(* CODESYS project BODAS_RC18-12_27-18_40.library
   DocFormat: reStructuredText
   Company: Bosch Rexroth AG
   DefaultNamespace: BODAS_RC18-12_27-18_40
   Title: BODAS_RC18-12_27-18_40
   Description: User library to use BODAS-BSW services (API) for RC40.
   Version: 3.0.1

Project tree, tasks and I/O mapping:
  Communication API/
    CAN/
      STRUCTURE/
        data type bds_can_BufManage_ts
        data type bds_can_DataboxBufInfo_ts
        data type bds_can_DataboxData08_ts
        data type bds_can_Message_ts
        data type bds_can_DataboxData64_ts
        data type bds_can_RxDatabox_ts
        data type bds_can_DataboxData_ts
        data type bds_can_TxDatabox_ts
      ENUM/
        data type bds_can_Chnl_te
      CAN legacy/
        API/
          function bds_can_getData [ST]
          function bds_can_getDatabox [ST]
          function bds_can_getRxBufStatus [ST]
          function bds_can_getStatus [ST]
          function bds_can_getTxBufStatus [ST]
          function bds_can_init [ST]
          function bds_can_initRxDatabox [ST]
          function bds_can_initTxDatabox [ST]
          function bds_can_initxt [ST]
          function bds_can_isTxChannelFree [ST]
          function bds_can_isTxDataboxFree [ST]
          function bds_can_sendData [ST]
          function bds_can_sendDatabox [ST]
          function bds_can_registerBusOffCallback [ST]
          function bds_can_setTxDelay [ST]
          function bds_can_start [ST]
          function bds_can_resetTxBuf [ST]
          function bds_can_stop [ST]
          function bds_can_registerRxCallback [ST]
      CAN signal based/
        API/
          function bds_can_sendSignal [ST]
          function bds_can_sendSignalGroup [ST]
          function bds_can_receiveSignal [ST]
          function bds_can_receiveSignalGroup [ST]
          function bds_can_setGroupSignalData [ST]
          function bds_can_setMsgGroup [ST]
          function bds_can_resetAllMsgGroups [ST]
          function bds_can_startAllMsgGroups [ST]
      UNION/
        data type bds_can_DataboxData_tu
      GVL/
        global variables GVL_can
      CAN_FFI_API/
        function bds_can_sendData_ffi [ST]
        function bds_can_getData_ffi [ST]
        function bds_can_getStatus_ffi [ST]
        function bds_can_isTxChannelFree_ffi [ST]
        function bds_can_getRxBufStatus_ffi [ST]
        function bds_can_getTxBufStatus_ffi [ST]
        function bds_can_sendDatabox_ffi [ST]
        function bds_can_getDatabox_ffi [ST]
        function bds_can_isTxDataboxFree_ffi [ST]
      CAN-FD legacy/
        API/
          function bds_can_fd_getData [ST]
          function bds_can_fd_getRxBufStatus [ST]
          function bds_can_fd_getTxBufStatus [ST]
          function bds_can_fd_isTxChannelFree [ST]
          function bds_can_fd_registerRxBuf [ST]
          function bds_can_fd_registerTxBuf [ST]
          function bds_can_fd_resetTxBuf [ST]
          function bds_can_fd_sendData [ST]
          function bds_can_fd_registerRxCallback [ST]
          function bds_can_fd_registerRxDataboxes [ST]
          function bds_can_fd_registerTxDataboxes [ST]
          function bds_can_fd_initRxDatabox [ST]
          function bds_can_fd_initTxDatabox [ST]
          function bds_can_fd_getDatabox [ST]
          function bds_can_fd_sendDatabox [ST]
          function bds_can_fd_isTxDataboxFree [ST]
          function bds_can_fd_setTxDelay [ST]
        ENUM/
          data type bds_can_fd_St_te
        STRUCTURE/
          data type bds_can_fd_Message_ts
          data type bds_can_fd_RxDatabox_ts
          data type bds_can_fd_DataboxData_ts
          data type bds_can_fd_DataboxBufInfo_ts
          data type bds_can_fd_BufManage_ts
          data type bds_can_fd_TxDatabox_ts
      CAN_FD_FFI_API/
        function bds_can_fd_getRxBufStatus_ffi [ST]
        function bds_can_fd_sendData_ffi [ST]
        function bds_can_fd_getTxBufStatus_ffi [ST]
        function bds_can_fd_getData_ffi [ST]
        function bds_can_fd_isTxChannelFree_ffi [ST]
        function bds_can_fd_getDatabox_ffi [ST]
        function bds_can_fd_sendDatabox_ffi [ST]
        function bds_can_fd_isTxDataboxFree_ffi [ST]
    ISOBUS/
      STRUCTURE/
        data type bds_isobus_appInst_ts
        data type bds_isobus_bamCtrl_ts
        data type bds_isobus_caName_ts
        data type bds_isobus_canID_ts
        data type bds_isobus_dtcList_ts
        data type bds_isobus_dtc_ts
        data type bds_isobus_err_ts
        data type bds_isobus_rxDataboxInfo_ts
        data type bds_isobus_rxEtpCtrl_ts
        data type bds_isobus_rxMsg_ts
        data type bds_isobus_rxTpCtrl_ts
        data type bds_isobus_txDataboxInfo_ts
        data type bds_isobus_txEtpCtrl_ts
        data type bds_isobus_txMsg_ts
        data type bds_isobus_txTpCtrl_ts
        data type bds_isobus_lamp_ts
        data type bds_isobus_nm_ts
        data type bds_isobus_aperiodicDataboxNum_ts
        data type bds_isobus_periodicDataboxNum_ts
        data type bds_isobus_caAddrInfoTbl_ts
        data type bds_isobus_caAddrInfoTblRef_ts
      UNION/
        data type bds_isobus_caName_tu
        data type bds_isobus_canID_tu
      API/
        function bds_isobus_cfgAddrClaimFormat [ST]
        function bds_isobus_getCaAddr [ST]
        isobus dtclist bds_isobus_getDiagnostic [ST]
        function bds_isobus_getRxDataboxStatus [ST]
        function bds_isobus_getStatus [ST]
        function bds_isobus_initComm [ST]
        isobus dtclist bds_isobus_initDiagnostic [ST]
        function bds_isobus_registerErrClrCbk [ST]
        function bds_isobus_registerInstances [ST]
        function bds_isobus_registerRxDataboxes [ST]
        function bds_isobus_registerTxDataboxes [ST]
        function bds_isobus_sendDatabox [ST]
        function bds_isobus_sendRequestPGN [ST]
        function bds_isobus_setCaAddr [ST]
        function bds_isobus_setCaInfo [ST]
        function bds_isobus_setCaName [ST]
        function bds_isobus_initFailureList [ST]
        function bds_isobus_initRxDatabox [ST]
        function bds_isobus_initTxDatabox [ST]
        function bds_isobus_registerCaAddrTable [ST]
        function bds_isobus_registerCaAddrInfoCbk [ST]
        function bds_isobus_getCaAddrByName [ST]
        function bds_isobus_getAddressInfoTblRecordSize [ST]
      GVL/
        global variables GVL_isobus
      J1939-76/
        STRUCTURE/
          data type bds_isobus_cnsrDataboxInfo_ts
          data type bds_isobus_cnsrSdgMsg_ts
          data type bds_isobus_cnsrSdgSeqNum_ts
          data type bds_isobus_prodDataboxInfo_ts
          data type bds_isobus_prodSdgMsg_ts
          data type bds_isobus_sftyTmr_ts
          data type bds_isobus_sfty_canID_ts
          data type bds_isobus_shmMsg_ts
        API/
          function bds_isobus_initCnsrSdgDatabox [ST]
          function bds_isobus_initProdSdgDatabox [ST]
          function bds_isobus_registerCnsrSdgDataboxes [ST]
          function bds_isobus_registerProdSdgDataboxes [ST]
        UNION/
          data type bds_isobus_sdmCrcVal_tu
          data type bds_isobus_sfty_canID_tu
        ENUM/
          data type bds_isobus_sdgCnsrStatus_te
          data type bds_isobus_sdgState_te
          data type bds_isobus_sfty_apiRetVal_te
      ENUM/
        data type bds_isobus_caAddrCbEventType_te
    LIN/
      API/
        function bds_lin_getStatus [ST]
        function bds_lin_gotoSleep [ST]
        function bds_lin_receiveSignal [ST]
        function bds_lin_sendSignal [ST]
        function bds_lin_setSchedule [ST]
        function bds_lin_wakeUp [ST]
      GVL/
        global variables GVL_lin
    Ethernet/
      API/
        function bds_ethIPv4_setLocalIpAdr [ST]
        function bds_ethIPv4_getLocalIpAdr [ST]
        function bds_ethIPv4_setDoipAdr [ST]
        function bds_ethIPv4_getLinkState [ST]
      STRUCTURE/
        data type bds_ethIPv4_getLocalIpAdr_ts
        data type bds_ethIPv4_setLocalIpAdr_ts
        data type bds_ethIPv4_LocalIpAdr_ts
        data type bds_ethIPv4_linkStateInfo_ts
      ENUMS/
        data type bds_ethIPv4_statusApi_te
        data type bds_ethIPv4_linkState_te
        data type bds_ethIPv4_retDoipAdr_te
        data type bds_ethIPv4_retLinkState_te
  Diagnostics API/
    UDS/
      API/
        function bds_uds_disable [ST]
        function bds_uds_GetActiveDid [ST]
        function bds_uds_getActiveSession [ST]
        function bds_uds_getNodeID [ST]
        function bds_uds_permitAccess [ST]
        function bds_uds_registerDidReadCallback [ST]
        function bds_uds_registerDidWriteCallback [ST]
        function bds_uds_registerRoutineCtrlCallback [ST]
        function bds_uds_registerRoutineF000Callback [ST]
        function bds_uds_setCallbackStatus [ST]
        function bds_uds_setUUID [ST]
        function bds_uds_updNodeIDinNVM [ST]
        function bds_uds_registerEvalKeyCallback [ST]
        function bds_uds_registerGetSeedCallback [ST]
        function bds_uds_registerRoutineF001Callback [ST]
        Vehicle Identification Number(VIN) APIs/
          function bds_uds_setVin [ST]
          function bds_uds_getVin [ST]
          function bds_uds_registerVinCallback [ST]
        function bds_uds_getActiveService [ST]
        function bds_uds_setNodeIdTesterId [ST]
      UNION/
        data type bds_uds_udsconfigparameter_tu
      STRUCTURE/
        data type bds_uds_udsconfigparameter_ts
        data type bds_uds_getActiveService_ts
      GVL/
        global variables GVL_uds
      FFI_API/
        function bds_uds_getActiveSession_ffi [ST]
        function bds_uds_getNodeID_ffi [ST]
        function bds_uds_getActiveService_ffi [ST]
        function bds_uds_getActiveDid_ffi [ST]
      ENUM/
        data type bds_udsCmn_statusApi_te
        data type bds_uds_setNodeIdTesterId_te
    XCP/
      API/
        function bds_xcp_setMode [ST]
      GVL/
        global variables GVL_xcp
  I/O API/
    SAFOUT/
      STRUCTURE/
        data type bds_safout_ts
      API/
        function bds_safout_resetError [ST]
        function bds_safout_ignoreError [ST]
        function bds_safout_getStatus [ST]
        function bds_safout_unlock [ST]
        function bds_safout [ST]
        function bds_safout_cfg [ST]
        function bds_safout_cfgDiag [ST]
        function bds_safout_enableTest [ST]
      GVL/
        global variables GVL_safout
    IN legacy/
      STRUCTURE/
        data type bds_in_aic_ts
        data type bds_in_fi_ts
        data type bds_in_FrqBuffered_ts
        data type bds_in_aiv_ts
        data type bds_in_sent_SDDataBox_ts
        data type bds_in_sent_slowData_ts
        data type bds_in_stPhase_ts
        data type bds_in_ri_ts
        data type bds_in_sent_BufManage_ts
        data type bds_in_sent_copyFDBuf_ts
        data type bds_in_sent_databoxinfo_ts
        data type bds_in_sent_decodedFD_ts
        data type bds_in_sent_FDBufInfo_ts
        data type bds_in_phase_ts
      API/
        function bds_in_aic_getStatus [ST]
        function bds_in_aid [ST]
        function bds_in_aid_cfg [ST]
        function bds_in_aiv [ST]
        function bds_in_aiv_cfg [ST]
        function bds_in_phase [ST]
        function bds_in_fi_cfg [ST]
        function bds_in_fi_getStatus [ST]
        function bds_in_phase_getStatus [ST]
        function bds_in_phase_resetCounter [ST]
        function bds_in_ri_cfg [ST]
        function bds_in_ri_cfgTemp [ST]
        function bds_in_sent_getSDDatabox [ST]
        function bds_in_sent_getStatus [ST]
        function bds_in_sent_initSDDatabox [ST]
        function bds_in_sent_registerCopyFDFifo [ST]
        function bds_in_sent_registerFDFifo [ST]
        function bds_in_ri_getStatus [ST]
        function bds_in_aiv_getStatus [ST]
        function bds_in_sent_registerSDDataboxes [ST]
        function bds_in_sent_getSD [ST]
        function bds_in_ri [ST]
        function bds_in_ai [ST]
        function bds_in_aic [ST]
        function bds_in_ri_getTemp [ST]
        function bds_in_sent_copyFDFifo [ST]
        function bds_in_sent_disable [ST]
        function bds_in_sent_enable [ST]
        function bds_in_sent_getFD [ST]
        function bds_in_aic_cfg [ST]
        function bds_in_di [ST]
        function bds_in_fi [ST]
        function bds_in_fi_buffered [ST]
      GVL/
        global variables GVL_in
    OUT_LEGACY/
      function bds_out_do_resetError [ST]
      function bds_out_do_unlock [ST]
      function bds_out_po [ST]
      function bds_out_poc [ST]
      function bds_out_poc_cfgDither [ST]
      function bds_out_poc_cfgPI [ST]
      function bds_out_po_cfgPwrLs [ST]
      function bds_out_po_cfg [ST]
      function bds_out_po_disableTstPls [ST]
      function bds_out_po_getCurrent [ST]
      function bds_out_po_getStatus [ST]
      function bds_out_po_resetError [ST]
      function bds_out_po_cfgPeriod [ST]
      function bds_out_po_disable [ST]
      function bds_out_aov_cfg [ST]
      function bds_out_aov_cfgPI [ST]
      function bds_out_aov_getStatus [ST]
      function bds_out_aov_getVoltage [ST]
      function bds_out_aov_resetError [ST]
      function bds_out_cfgLoadCharacteristic [ST]
      function bds_out_do [ST]
      function bds_out_do_cfgPwrLs [ST]
      function bds_out_do_disable [ST]
      function bds_out_aov [ST]
      function bds_out_do_disableTstPls [ST]
      function bds_out_do_getCurrent [ST]
      function bds_out_pod [ST]
      function bds_out_do_getStatus [ST]
      function bds_out_poc_cfg [ST]
      function bds_out_po_unlock [ST]
    OUT/
      API/
        function bds_outClcU_setVoltage [ST]
        function bds_outClcU_setPercUBat [ST]
        function bds_outClcU_get [ST]
        function bds_outClcU_rstErr [ST]
        function bds_outDig_set [ST]
        function bds_outDig_get [ST]
        function bds_outDig_cfgDiag [ST]
        function bds_outDig_rstErr [ST]
        function bds_outPwm_setDutyCycle [ST]
        function bds_outPwm_get [ST]
        function bds_outPwm_cfgPeriod [ST]
        function bds_outPwm_rstErr [ST]
        function bds_outPwm_cfgDiag [ST]
        function bds_outPwm_cfgMode [ST]
        function bds_outPwm_setCurrent [ST]
        function bds_outPwm_cfgDiagCurrentDe [ST]
        function bds_outPwm_cfgClc [ST]
        function bds_outPwm_cfgDither [ST]
        function bds_outClcU_cfgClc [ST]
      STRUCTURE/
        data type bds_out_do_ts
        data type bds_out_po_ts
        data type bds_out_aov_ts
        data type bds_outClcU_setVoltage_ts
        data type bds_outClcU_setPercUBat_ts
        data type bds_outClcU_get_ts
        data type bds_outCmn_statusDiag_tb
        data type bds_outClcU_rstErr_ts
        data type bds_outDig_set_ts
        data type bds_outDig_get_ts
        data type bds_outDig_cfgDiag_ts
        data type bds_outDig_rstErr_ts
        data type bds_outPwm_setDutyCycle_ts
        data type bds_outPwm_get_ts
        data type bds_outPwm_cfgPeriod_ts
        data type bds_outPwm_rstErr_ts
        data type bds_outPwm_cfgDiag_ts
        data type bds_outPwm_cfgMode_ts
        data type bds_outPwm_setCurrent_ts
        data type bds_outPwm_cfgDiagCurrentDe_ts
        data type bds_outPwm_cfgDither_ts
        data type bds_outClcU_cfgClc_ts
        data type bds_outClcU_clcParams_ts
        data type bds_outCmn_diagParam_ts
        data type bds_outPwm_cfgClc_ts
        data type bds_outPwm_clcParams_ts
        data type bds_outPwm_ditherParams_ts
      ENUM/
        data type bds_load_characteristic_te
        data type bds_outCmn_statusApi_te
        data type bds_outPwm_cfgMode_te
        data type bds_outPwm_cfgDither_te
      GVL/
        global variables GVL_out
      FFI_API/
        function bds_out_aov_ffi [ST]
        function bds_out_aov_cfg_ffi [ST]
        function bds_out_aov_cfgPI_ffi [ST]
        function bds_out_aov_getStatus_ffi [ST]
        function bds_out_aov_getVoltage_ffi [ST]
        function bds_out_cfgLoadCharacteristic_ffi [ST]
        function bds_out_do_ffi [ST]
        function bds_out_do_cfgPwrLs_ffi [ST]
        function bds_out_do_disable_ffi [ST]
        function bds_out_do_disableTstPls_ffi [ST]
        function bds_out_do_getCurrent_ffi [ST]
        function bds_out_do_getStatus_ffi [ST]
        function bds_out_po_ffi [ST]
        function bds_out_poc_ffi [ST]
        function bds_out_poc_cfg_ffi [ST]
        function bds_out_poc_cfgDither_ffi [ST]
        function bds_out_poc_cfgPI_ffi [ST]
        function bds_out_pod_ffi [ST]
        function bds_out_po_cfg_ffi [ST]
        function bds_out_po_cfgPeriod_ffi [ST]
        function bds_out_po_cfgPwrLs_ffi [ST]
        function bds_out_po_disable_ffi [ST]
        function bds_out_po_disableTstPls_ffi [ST]
        function bds_out_po_getCurrent_ffi [ST]
        function bds_out_po_getStatus_ffi [ST]
    SENT/
      STRUCTURE/
        data type bds_sent_chSt_tb
        data type bds_sent_rxFastData_ts
        data type bds_sent_rxSlowData_ts
        data type bds_sent_getSlowDataBufd_ts
        data type bds_sent_getFastDataBufd_ts
        data type bds_sent_fastDataMsg_ts
        data type bds_sent_fastDataBuf_ts
        data type bds_sent_slowDataMsg_ts
        data type bds_sent_slowDataBuf_ts
      ENUM/
        data type bds_sentCmn_status_te
      API/
        function bds_sent_getFastData [ST]
        function bds_sent_getSlowData [ST]
        function bds_sent_getFastDataBufd [ST]
        function bds_sent_getSlowDataBufd [ST]
      FFI_API/
        function bds_sent_getFastData_ffi [ST]
        function bds_sent_getFastDataBufd_ffi [ST]
        function bds_sent_getSlowData_ffi [ST]
        function bds_sent_getSlowDataBufd_ffi [ST]
    IN/
      STRUCTURE/
        data type bds_inI_measmt_ts
        data type bds_inDig_measmt_ts
        data type bds_inCmn_pullParam_ts
        data type bds_inI_cfgPull_ts
        data type bds_inI_shunt_ts
        data type bds_inDig_cfgPull_ts
        data type bds_inPwm_tiMeasmt_ts
        data type bds_inPwm_tiBufdMeasmt_ts
        data type bds_inPwm_frqMeasmt_ts
        data type bds_inPwm_tiBufd_ts
        data type bds_inR_measmt_ts
        data type bds_inU_measmt_ts
        data type bds_inU_cfgPull_ts
        data type bds_inPha_measmt_ts
        data type bds_inPha_statusDiag_tb
        data type bds_inPha_tiBufdMeasmt_ts
        data type bds_inPha_tiBufd_ts
      ENUM/
        data type bds_inCmn_status_te
        data type bds_inCmn_pullType_te
        data type bds_inI_stShunt_te
        data type bds_inCmn_iPull_te
      API/
        function bds_inI_cfgPull [ST]
        function bds_inI_ctrlShunt [ST]
        function bds_inDig_get [ST]
        function bds_inI_get [ST]
        function bds_inDig_cfgPull [ST]
        function bds_inPwm_getTi [ST]
        function bds_inPwm_getTiBufd [ST]
        function bds_inR_get [ST]
        function bds_inPwm_getFrq [ST]
        function bds_inU_get [ST]
        function bds_inU_cfgPull [ST]
        function bds_inPha_get [ST]
        function bds_inPha_getTiBufd [ST]
      FFI_API/
        function bds_inDig_cfgPull_ffi [ST]
        function bds_inI_cfgPull_ffi [ST]
        function bds_inI_ctrlShunt_ffi [ST]
        function bds_inPwm_getFrq_ffi [ST]
        function bds_inPwm_getTi_ffi [ST]
        function bds_inPwm_getTiBufd_ffi [ST]
        function bds_inU_cfgPull_ffi [ST]
  Memory API/
    NVM/
      API/
        function bds_mem_getBlockStatus [ST]
        function bds_mem_markBlock [ST]
        function bds_mem_readBlock [ST]
        function bds_mem_writeBlock [ST]
      GVL/
        global variables GVL_mem
      FFI_API/
        function bds_mem_getBlockStatus_ffi [ST]
        function bds_mem_markBlock_ffi [ST]
        function bds_mem_readBlock_ffi [ST]
        function bds_mem_writeBlock_ffi [ST]
  System API/
    SEC/
      ENUM/
        data type bds_diag_inst_te
        data type bds_sec_securityOperations_te
      API/
        function bds_sec_evalRespKey [ST]
        function bds_sec_getLevel [ST]
        function bds_sec_getRnd [ST]
        function bds_sec_resetLevel [ST]
        function bds_sec_saveSecret [ST]
        function bds_sec_scrambleRexrothSecretsPerm [ST]
        function bds_sec_setLevel [ST]
        function bds_sec_getSeed [ST]
      GVL/
        global variables GVL_sec
    SYS/
      API/
        function bds_sys_ait [ST]
        function bds_sys_aiv [ST]
        function bds_sys_cancelAltWakeup [ST]
        function bds_sys_di [ST]
        function bds_sys_do [ST]
        function bds_sys_getAge [ST]
        function bds_sys_getCoreLoad [ST]
        function bds_sys_getEcuInfo [ST]
        function bds_sys_getResetInfo [ST]
        function bds_sys_getStates [ST]
        function bds_sys_getT15 [ST]
        function bds_sys_getTaskRuntime [ST]
        function bds_sys_getTime [ST]
        function bds_sys_getVersion [ST]
        function bds_sys_getVSS [ST]
        function BDS_SYS_GET_LOCK_COMMON [ST]
        function bds_sys_memByteCopy [ST]
        function bds_sys_releasePostRunProlong [ST]
        function BDS_SYS_RELEASE_LOCK_COMMON [ST]
        function bds_sys_requestPostRunProlong [ST]
        function bds_sys_resetCoreLoad [ST]
        function bds_sys_resetEcu [ST]
        function bds_sys_resetINH [ST]
        function bds_sys_setVSS [ST]
        function bds_sys_startLoader [ST]
        function bds_sysPb_getVariant [ST]
        function bds_sysPb_cfgVariant [ST]
        function bds_sys_applSwName [ST]
        function bds_sysSm_getCfg [ST]
        function bds_sys_regOverwriteOpHrsCbk [ST]
        function bds_codesys_setForcingWritingMode [ST]
      ENUM/
        data type bds_sys_coreid_te
        data type bds_sys_states_te
        data type bds_sys_task_te
        data type bds_sysCmn_status_te
        data type bds_sys_aswNameStatus_te
        data type bds_sys_regOverwriteOpHrs_te
      STRUCTURE/
        data type bds_sys_coreload_info_ts
        data type bds_sys_states_ts
        data type bds_sys_taskruntime_ts
        data type bds_ResetInfo_ts
        data type bds_EcuInfo_ts
        data type bds_sysPb_retValCfgVrnt_ts
        data type bds_sysPb_vrntParam_ts
        data type bds_sysPb_retValGetVrnt_ts
        data type bds_sys_retValApplSwName_ts
      GVL/
        global variables GVL_sys
      FFI_API/
        function bds_sysPb_getVariant_ffi [ST]
        function bds_sys_getAge_ffi [ST]
        function bds_sys_getCoreLoad_ffi [ST]
        function bds_sys_getEcuInfo_ffi [ST]
        function bds_sys_getResetInfo_ffi [ST]
        function bds_sys_getStates_ffi [ST]
        function bds_sys_getTaskRuntime_ffi [ST]
        function bds_sys_getTime_ffi [ST]
        function bds_sys_getVersion_ffi [ST]
    DSM/
      STRUCTURE/
        data type bds_dfes_ts
        data type bds_dsm_j1939Lamp_ts
        data type bds_dsm_J1939_info_ts
        data type bds_dsm_dfc_ts
        data type bds_dsm_dtcj1939_ts
        data type bds_dsm_fid_ts
      API/
        function bds_dsm_delError [ST]
        function bds_dsm_delErrors [ST]
        function bds_dsm_delErrorsJ1939 [ST]
        function bds_dsm_delError_DTC [ST]
        Macro Functions/
          function bds_dsm_DFC_da [ST]
          function bds_dsm_DFC_dfl [ST]
          function bds_dsm_DFC_fl [ST]
          function bds_dsm_DFC_fsc [ST]
          function bds_dsm_DFC_ldf [ST]
          function bds_dsm_DFC_ms [ST]
          function bds_dsm_DFC_t [ST]
          function bds_dsm_DFC_tf [ST]
          function bds_dsm_DFC_tsc [ST]
        function bds_dsm_getErrors [ST]
        function bds_dsm_getDTC_Status [ST]
        function bds_dsm_getErrors_DTC [ST]
        function bds_dsm_getFIdPermission [ST]
        function bds_dsm_getNumErrors [ST]
        function bds_dsm_getNumErrorsJ1939 [ST]
        function bds_dsm_testError [ST]
        function bds_dsm_test_ErrorDFC [ST]
        function bds_dsm_test_ErrorDTC [ST]
        function bds_dsm_updateDebError [ST]
        function bds_dsm_updateError [ST]
        function bds_dsm_updateError_DTC [ST]
        function bds_dsm_getDFC_Status [ST]
        function bds_dsm_getDFES [ST]
        function bds_dsm_getErrorsJ1939 [ST]
        function bds_dsm_getDFES_DTC [ST]
        function bds_dsm_getDTC_DFC [ST]
        function bds_dsm_getDTC_DFCJ1939 [ST]
        function bds_dsm_getDTC_J1939 [ST]
      ENUM/
        data type bds_dsm_state_te
      GVL/
        global variables GVL_dsm
      FFI_API/
        function bds_dsm_getErrors_ffi [ST]
        function bds_dsm_updateError_ffi [ST]
        function bds_dsm_getNumErrors_ffi [ST]
        function bds_dsm_getDFC_Status_ffi [ST]
      DSM Refactored( 3-byte DTC)/
        STRUCTURE/
          data type bds_dsmCmn_stWord_tb
          data type bds_dsmDTC_deleteErr_ts
          data type bds_dsmDTC_getDFES_ts
          data type bds_dsmDTC_getDTCVal_ts
          data type bds_dsmDTC_getErrList_ts
          data type bds_dsmDTC_getStatus_ts
          data type bds_dsmDTC_updateErr_ts
          data type bds_dsmJ1939_LampSt_tb
          data type bds_dsmJ1939_getJ1939DTC_ts
        API/
          function bds_dsmDTC_getDTCVal [ST]
          function bds_dsmDTC_updateErr [ST]
          function bds_dsmDTC_deleteErr [ST]
          function bds_dsmDTC_getErrList [ST]
          function bds_dsmDTC_getStatus [ST]
          function bds_dsmDTC_getDFES [ST]
          function bds_dsmJ1939_getJ1939DTC [ST]
        ENUM/
          data type bds_dsmCmn_st_te
          data type bds_dsmCmn_errState_te
          data type bds_dsmCmn_fltLvl_te
*)

// Communication API/CAN/STRUCTURE/bds_can_BufManage_ts
{attribute 'external_name' := 'cmp_rts_bds_can_BufManage_ts'}
TYPE bds_can_BufManage_ts :
STRUCT
	length_u16: UINT;
	idx_in_u16: UINT;
	idx_out_u16: UINT;
	BufEmpty_l: BOOL;
	BufOvfl_l: BOOL;
END_STRUCT
END_TYPE

// Communication API/CAN/ENUM/bds_can_Chnl_te
{attribute 'external_name' := 'cmp_rts_bds_can_Chnl_te'}
TYPE bds_can_Chnl_te :
(
	///CAN channel 1
	BDS_CAN_1_D := 0,
	///CAN channel 2
	BDS_CAN_2_D,
	///CAN channel 3
	BDS_CAN_3_D,
	///CAN channel 4
	BDS_CAN_4_D,
	BDS_CAN_NBR_E
)USINT;
END_TYPE

// Communication API/CAN/STRUCTURE/bds_can_DataboxBufInfo_ts
{attribute 'external_name' := 'cmp_rts_bds_can_DataboxBufInfo_ts'}
TYPE bds_can_DataboxBufInfo_ts :
STRUCT
	start_pas: POINTER TO bds_can_DataboxData_ts;
	Manage_s: bds_can_BufManage_ts;
END_STRUCT
END_TYPE

// Communication API/CAN/STRUCTURE/bds_can_DataboxData08_ts
{attribute 'external_name' := 'cmp_rts_bds_can_DataboxData08_ts'}
TYPE bds_can_DataboxData08_ts :
STRUCT
	data_au8: ARRAY[0..7] OF USINT;
	numBytes_u8: USINT;
END_STRUCT
END_TYPE

// Communication API/CAN/UNION/bds_can_DataboxData_tu
{attribute 'external_name' := 'cmp_rts_bds_can_DataboxData_tu'}
TYPE bds_can_DataboxData_tu :

UNION
	len08_s: bds_can_DataboxData08_ts;
	len64_s: bds_can_DataboxData64_ts;
END_UNION

END_TYPE

// Communication API/CAN/STRUCTURE/bds_can_Message_ts
{attribute 'external_name' := 'cmp_rts_bds_can_Message_ts'}
TYPE bds_can_Message_ts :
STRUCT
	///Identifier of the message.
	id_u32: UDINT;
	///Format which will be transmitted (Standard / Extended)
	format_u8: USINT;
	///Number of data bytes which will be transmitted or which where received.
	numBytes_u8: USINT;
	///Data which will be transmitted or which were received.
	data_au8: ARRAY[0..7] OF USINT;
END_STRUCT
END_TYPE

// Communication API/CAN/STRUCTURE/bds_can_DataboxData64_ts
{attribute 'external_name' := 'cmp_rts_bds_can_DataboxData64_ts'}
TYPE bds_can_DataboxData64_ts :
STRUCT
	data_au8: ARRAY[0..63] OF USINT;
	numBytes_u8: USINT;
END_STRUCT
END_TYPE

// Communication API/CAN/STRUCTURE/bds_can_RxDatabox_ts
{attribute 'external_name' := 'cmp_rts_bds_can_RxDatabox_ts'}
TYPE bds_can_RxDatabox_ts :
STRUCT
	id_u32: UDINT;
	format_u8: USINT;
	numBytes_u8: USINT;
	callback_pf: UDINT;
	Buf_s: bds_can_DataboxBufInfo_ts;
END_STRUCT
END_TYPE

// Communication API/CAN/STRUCTURE/bds_can_DataboxData_ts
{attribute 'external_name' := 'cmp_rts_bds_can_DataboxData_ts'}
TYPE bds_can_DataboxData_ts :
STRUCT
	///Data which will be transmitted or which were received.
	data_au8: ARRAY[0..7] OF USINT;
	///Number of data bytes which will be transmitted or which where received.
	numBytes_u8: USINT;
END_STRUCT
END_TYPE

// System API/DSM/STRUCTURE/bds_dfes_ts
{attribute 'external_name' := 'cmp_rts_bds_dfes_ts'}
TYPE bds_dfes_ts :
STRUCT
	/// REFERENCE number
	id: UINT := 12;
	/// assigned predebouncing mode
	debmode: UINT := 4;
END_STRUCT
END_TYPE

// System API/SEC/ENUM/bds_diag_inst_te
{attribute 'external_name' := 'cmp_rts_bds_diag_inst_te'}
TYPE bds_diag_inst_te :
(
	BDS_SEC_ASW_START_INSTANCE_E := 0,
	BDS_SEC_ASW_INST_NAME_1_E := BDS_SEC_ASW_START_INSTANCE_E,
	BDS_SEC_ASW_INST_NAME_2_E,
	BDS_SEC_ASW_INST_NAME_3_E,
	BDS_SEC_ASW_NUM_INSTANCE_E
);
END_TYPE

// I/O API/OUT/STRUCTURE/bds_out_do_ts
{attribute 'external_name' := 'cmp_rts_bds_out_do_ts'}
TYPE bds_out_do_ts :
STRUCT
	///status flags for status_b16 
	///	initOut_DB16: USINT := 16#1;(*initialization after startup*)
	///	
	///	cfgPOC_DB16: USINT := 16#2;(*configuration of closed loop control*)
	///	
	///	cfgPeriod_DB16: USINT := 16#4;(*configuration of period*)
	///	
	///	cfgDither_DB16: USINT := 16#8;(*configuration of dither*)
	///	
	///	cfgDeviation_DB16: USINT := 16#10;(*configuration of deviation*)
	///	
	///	cfgPI_DB16: USINT := 16#20;(*configuration of KpKi*)
	///	
	///	lockedSCB_DB16: USINT := 16#40;(*locked by SCB...necessary for AOV*)
	///	
	///	lockedSCG_DB16: USINT := 16#80;(*locked by SCG...necessary for AOV*)
	///	
	///	lockedOC_DB16: UINT := 16#100;(*locked by OC*)
	///	
	///	locked_DB16: UINT := 16#200;(*locked by Error Handler*)
	///	
	///	lockedMO_DB16: UINT := 16#400;(*locked by Monitoring Module (MO) Error*)
	///	
	///	lockCouTiReact_DB16: UINT := 16#800;(*locked reactivation timer reload after a hot short circuit*)
	///	
	///	tiReactNotElapsed_DB16: UINT := 16#1000;(*time for reactivation after a hot short circuit not elapsed*)
	///	
	///	linked_DB16: UINT := 16#2000;(*linked at least with one other safout output*)
	///	
	///	tlsPlsDis_DB16: UINT:=16#4000;(*Test pulses disable*)
	///	
	///	disabled_DB16: UINT := 16#8000;(*output is disabled (avoid open load faults of unused outputs)*)
	///	
	///	cfgOutMask_DB16: UINT := ((((cfgPI_DB16 OR cfgDeviation_DB16) OR cfgDither_DB16) OR cfgPeriod_DB16) OR cfgPOC_DB16);
	status_b16: UINT;
	///state
	state_u8: USINT;
	///ADC digits, range from 0..25000
	digits_u16: UINT;
	///actual current [mA]
	iAct_u16: UINT;
	///fault status
	stDFC_SCB_u16: UINT;
	///fault status
	stDFC_SCG_u16: UINT;
	///fault status
	stDFC_OL_u16: UINT;
	///fault status
	stDFC_OT_u16: UINT;
	///fault status
	stDFC_OC_u16: UINT;
	///Unintended switch ON of output
	unintendedSwitchONErr_l: BOOL;
	///locked by Inhibits
	lockedByINH_l: BOOL;
END_STRUCT
END_TYPE

// I/O API/IN legacy/STRUCTURE/bds_in_aic_ts
{attribute 'external_name' := 'cmp_rts_bds_in_aic_ts'}
TYPE bds_in_aic_ts :
STRUCT
	///status flags for status_b16 
	///	
	///	initIn_DB16: USINT := 16#1;(*initialization after startup*)
	///	
	///	cfgAiv_DB16: USINT := 16#2;(*configured for AIV thresholds*)
	///	
	///	cfgAic_DB16: USINT := 16#4;(*configured for AIC thresholds*)
	///	
	///	cfgAid_DB16: USINT := 16#8;(*configured for AID thresholds*)
	///	
	///	cfgRi_DB16: USINT := 16#10;(*configured for RI thresholds*)
	///	
	///	cfgFreq_DB16: USINT := 16#20;(*configured for standard frequency sensor*)
	///	
	///	cfgFreqDSM_DB16: USINT := 16#40;(*configured for DSM frequency sensor*)
	///	
	///	lostSignalInfoDSM_DB16: USINT := 16#80;
	///	
	///	actShunt_DB16: UINT := 16#1000;(*shunt is activated for DSM sensor respective AIC*)
	///	
	///	lockReactShunt_DB16: UINT := 16#2000;(*locked shunt reactivation*)
	///	
	///	cfgInMask_DB16: UINT := (((((cfgFreqDSM_DB16 OR cfgFreq_DB16) OR cfgRi_DB16) OR cfgAid_DB16) OR cfgAic_DB16) OR cfgAiv_DB16);
	status_b16: UINT;
	///ADC digits, range from 0..25000
	digits_u16: UINT;
	///current [µA]
	i_uA_u16: UINT;
	///fault status
	stDFC_SCB_u16: UINT;
	///fault status
	stDFC_SCG_u16: UINT;
END_STRUCT
END_TYPE

// I/O API/IN legacy/STRUCTURE/bds_in_fi_ts
{attribute 'external_name' := 'cmp_rts_bds_in_fi_ts'}
TYPE bds_in_fi_ts :
STRUCT
	///status flags for status_b16 
	///	
	///	initIn_DB16: USINT := 16#1;(*initialization after startup*)
	///	
	///	cfgAiv_DB16: USINT := 16#2;(*configured for AIV thresholds*)
	///	
	///	cfgAic_DB16: USINT := 16#4;(*configured for AIC thresholds*)
	///	
	///	cfgAid_DB16: USINT := 16#8;(*configured for AID thresholds*)
	///	
	///	cfgRi_DB16: USINT := 16#10;(*configured for RI thresholds*)
	///	
	///	cfgFreq_DB16: USINT := 16#20;(*configured for standard frequency sensor*)
	///	
	///	cfgFreqDSM_DB16: USINT := 16#40;(*configured for DSM frequency sensor*)
	///	
	///	lostSignalInfoDSM_DB16: USINT := 16#80;
	///	
	///	actShunt_DB16: UINT := 16#1000;(*shunt is activated for DSM sensor respective AIC*)
	///	
	///	lockReactShunt_DB16: UINT := 16#2000;(*locked shunt reactivation*)
	///	
	///	cfgInMask_DB16: UINT := (((((cfgFreqDSM_DB16 OR cfgFreq_DB16) OR cfgRi_DB16) OR cfgAid_DB16) OR cfgAic_DB16) OR cfgAiv_DB16);
	///	
	///	standstill_DU8: USINT := 16#0;(*standstill*)
	///	
	///	dirLeft_DU8: USINT := 16#1;(*direction left*)
	///	
	///	dirRight_DU8: USINT := 16#2;(*direction right*)
	///	
	///	dirUnknown_DU8: USINT := 16#4;(*direction not known for sure (e.g. after standstill)*)
	///	
	///	noError_DU8: USINT := 16#0;(*error free*)
	///	
	///	airGapError_DU8: USINT := 16#1;(*air gap error (pulse is shorter than 64us)*)
	///	
	///	mountError_DU8: USINT := 16#2;(*mounting error (pulse is longer than 254us)*)
	///	
	///	signalLengthError_DU8: USINT := 16#4;(*undefined signal length - should not occur (pulse is longer than 1785us*)
	///	
	///	signalError_DU8: USINT := 16#8;(*period too long or measured period exceeds maximum period*)
	///	
	///	noStatusAvailable_DU8: USINT := 16#10;(*no status signal available (frequency to high)*)
	///	
	///	diagSCUBAT_DU8: USINT := 16#20;
	///	
	///	diagSCGND_OR_OL_DU8: USINT := 16#40;
	///	
	///	maskFrequency_DU32: UDINT := 16#FFFFF;(*DSM mask to get the frequency out*)
	///	
	///	maskDirection_DU32: UDINT := 16#F00000;(*DSM mask to get the direction*)
	///	
	///	numShiftDirection_DU32: USINT := 20;(*DSM shift number to get the direction*)
	///	
	///	maskStatus_DU32: UDINT := 16#FF000000;(*DSM mask to get the status*)
	///	
	///	numShiftStatus_DU32: USINT := 24;(*DSM shift number to get the status*)
	status_b16: UINT;
	///current dutycycle [100%=16#8000]
	rDutycycle_u32: UDINT;
	///last high_time duration [µs]
	tiPulse_u32: UDINT;
	///period duration [µs]
	tiPeriod_u32: UDINT;
	///signal period counter
	ctPeriod_u32: UDINT;
	///signal state
	///   + Bit0 state at function call time ("1" for high or "0" for low
	///   + Bit1 no update available (request within the same period)
	///   + Bit2 period too long (timer overflow)
	///   + Bit3 measured period exceeds given maximum length 
	stSignal_u8: USINT;
	///frequency in [dHz]
	f_dHz_u32: UDINT;
	///period duration [µs] for DSM sensor
	tiPeriodDSM_u32: UDINT;
	///frequency of DSM in [dHz] (see defines above)
	f_dHzDSM_u32: UDINT;
	///direction (see defines above)
	directionDSM_u8: USINT;
	///status
	statusDSM_u8: USINT;
END_STRUCT
END_TYPE

// I/O API/IN legacy/STRUCTURE/bds_in_FrqBuffered_ts
{attribute 'external_name' := 'cmp_rts_bds_in_FrqBuffered_ts'}
TYPE bds_in_FrqBuffered_ts :
STRUCT
	///Pointer of the start address of the period array
	tiPeriod_pu32: POINTER TO UDINT;
	///Pointer of the start address of the pulse array
	tiPulse_pu32: POINTER TO UDINT;
END_STRUCT
END_TYPE

// Communication API/CAN/STRUCTURE/bds_can_TxDatabox_ts
{attribute 'external_name' := 'cmp_rts_bds_can_TxDatabox_ts'}
TYPE bds_can_TxDatabox_ts :
STRUCT
	id_u32: UDINT;
	format_u8: USINT;
	numBytes_u8: USINT;
	data_au8: ARRAY[0..7] OF USINT;
	empty_l: BOOL;
	init_l: BOOL;
END_STRUCT
END_TYPE

// System API/SEC/ENUM/bds_sec_securityOperations_te
{attribute 'external_name' := 'cmp_rts_bds_sec_securityOperations_te'}
TYPE bds_sec_securityOperations_te :
(
	SEC_SRV_ReadDeviceInfo_E := 0,
	SEC_SRV_ChangePwdRexroth_E,
	SEC_SRV_ReadMemAddress_E,
	SEC_SRV_WriteMemAddress_E,
	SEC_SRV_StoreChangedDids_E,
	SEC_SRV_FlashBC_E,
	SEC_SRV_FlashCB_E,
	SEC_SRV_ChangeCustPwd_E,
	SEC_SRV_ReadDtc_E,
	SEC_SRV_ClearDtcCust_E,
	SEC_SRV_ClearDtcRexroth_E,
	SEC_SRV_ControlDtc_E,
	SEC_SRV_EcuReset_E
);
END_TYPE

// System API/SYS/ENUM/bds_sys_coreid_te
{attribute 'external_name' := 'cmp_rts_bds_sys_coreid_te'}
TYPE bds_sys_coreid_te :
(
	///ECU logical Core 0.
	BDS_CORE_0_D := 0,
	///ECU logical Core 1.
	BDS_CORE_1_D,
	///ECU logical Core 2.
	BDS_CORE_2_D,
	///ECU logical Core 3.
	BDS_CORE_3_D
)USINT;
END_TYPE

// System API/SYS/STRUCTURE/bds_sys_coreload_info_ts
{attribute 'external_name' := 'cmp_rts_bds_sys_coreload_info_ts'}
TYPE bds_sys_coreload_info_ts :
STRUCT
	///Core load of CPU.
	coreload_u16: UINT;
	///Maximum current cycle core load of CPU.
	coreload_max_currentcycle_u16: UINT;
	///Maximum life cycle core load of CPU.
	coreload_max_lifecycle_u16: UINT;
END_STRUCT
END_TYPE

// I/O API/SAFOUT/STRUCTURE/bds_safout_ts
{attribute 'external_name' := 'cmp_rts_bds_safout_ts'}
TYPE bds_safout_ts :
STRUCT
	/// channel (mode|number) 
	chnl_u16: UINT;
	/// status 
	status_b16: UINT;
	/// common state/setpoint 
	setOutCo_u16: UINT;
	/// partial state(s)/setpoint(s) 
	setOut1_u16: UINT;
	setOut2_u16: UINT;
	setOut3_u16: UINT;
	setOut4_u16: UINT;
	/// common current 
	iOutCo_u16: UINT;
	iOut1_u16: UINT;
	iOut2_u16: UINT;
	iOut3_u16: UINT;
	iOut4_u16: UINT;
	/// sum of the partial currents 
	iOutSum_u16: UINT;
	/// diagnostic info (summarized faults of the outputs) 
	diag_u32: UDINT;
	/// diagnostic info of previous cycle (not frozen) 
	diag2_u32: UDINT;
	/// channel is locked by output faults 
	stDFC_u16: UINT;
	/// channel is locked by current deviation fault 
	stDFC_iDev_u16: UINT;
	/// test status  
	testSts_u16: UINT;
END_STRUCT
END_TYPE

// System API/SYS/ENUM/bds_sys_states_te
{attribute 'external_name' := 'cmp_rts_bds_sys_states_te'}
TYPE bds_sys_states_te :
(
	///System is in initialization state.
	BDS_SYSSTATE_INIT_E := 0,
	///Initialization state is finished and cyclic tasks are running.
	BDS_SYSSTATE_RUN_E,
	///System is in Postrun state
	BDS_SYSSTATE_POSTRUN_E,
	///System is in shutdown state.
	BDS_SYSSTATE_SHUTDOWN_E
);
END_TYPE

// System API/SYS/STRUCTURE/bds_sys_states_ts
{attribute 'external_name' := 'cmp_rts_bds_sys_states_ts'}
TYPE bds_sys_states_ts :
STRUCT
	///Current state
	currentState_e: bds_sys_states_te;
	///Previous state
	prvState_e: bds_sys_states_te;
END_STRUCT
END_TYPE

// System API/SYS/STRUCTURE/bds_sys_taskruntime_ts
{attribute 'external_name' := 'cmp_rts_bds_sys_taskruntime_ts'}
TYPE bds_sys_taskruntime_ts :
STRUCT
	///Current net runtime.
	curr_net_runtime_u32: UDINT;
	///Maximum net runtime.
	max_net_runtime_u32: UDINT;
	///Minimum net runtime.
	min_net_runtime_u32: UDINT;
	///Average net runtime.
	avg_net_runtime_u32: UDINT;
	///Current gross runtime.
	curr_gross_runtime_u32: UDINT;
	///Maximum gross runtime.
	max_gross_runtime_u32: UDINT;
	///Minimum gross runtime.
	min_gross_runtime_u32: UDINT;
END_STRUCT
END_TYPE

// System API/SYS/ENUM/bds_sys_task_te
{attribute 'external_name' := 'cmp_rts_bds_sys_task_te'}
TYPE bds_sys_task_te :
(
	///100 ms cyclic task(low priority)
	Task_100ms_D := 0,
	///80 ms cyclic task
	Task_80ms_D,
	///50 ms cyclic task
	Task_50ms_D,
	///40 ms cyclic task
	Task_40ms_D,
	///20 ms cyclic task
	Task_20ms_D,
	///10 ms cyclic task
	Task_10ms_D,
	///5 ms cyclic task
	Task_5ms_D,
	///2 ms cyclic task
	Task_2ms_D,
	///1 ms cyclic task (high priority).
	Task_1ms_D
);
END_TYPE

// I/O API/OUT/STRUCTURE/bds_out_po_ts
{attribute 'external_name' := 'cmp_rts_bds_out_po_ts'}
TYPE bds_out_po_ts :
STRUCT
	///status flags for status_b16 
	///	initOut_DB16: USINT := 16#1;(*initialization after startup*)
	///	
	///	cfgPOC_DB16: USINT := 16#2;(*configuration of closed loop control*)
	///	
	///	cfgPeriod_DB16: USINT := 16#4;(*configuration of period*)
	///	
	///	cfgDither_DB16: USINT := 16#8;(*configuration of dither*)
	///	
	///	cfgDeviation_DB16: USINT := 16#10;(*configuration of deviation*)
	///	
	///	cfgPI_DB16: USINT := 16#20;(*configuration of KpKi*)
	///	
	///	lockedSCB_DB16: USINT := 16#40;(*locked by SCB...necessary for AOV*)
	///	
	///	lockedSCG_DB16: USINT := 16#80;(*locked by SCG...necessary for AOV*)
	///	
	///	lockedOC_DB16: UINT := 16#100;(*locked by OC*)
	///	
	///	locked_DB16: UINT := 16#200;(*locked by Error Handler*)
	///	
	///	lockedMO_DB16: UINT := 16#400;(*locked by Monitoring Module (MO) Error*)
	///	
	///	lockCouTiReact_DB16: UINT := 16#800;(*locked reactivation timer reload after a hot short circuit*)
	///	
	///	tiReactNotElapsed_DB16: UINT := 16#1000;(*time for reactivation after a hot short circuit not elapsed*)
	///	
	///	linked_DB16: UINT := 16#2000;(*linked at least with one other safout output*)
	///	
	///	tlsPlsDis_DB16: UINT:=16#4000;(*Test pulses disable*)
	///	
	///	disabled_DB16: UINT := 16#8000;(*output is disabled (avoid open load faults of unused outputs)*)
	///	
	///	cfgOutMask_DB16: UINT := ((((cfgPI_DB16 OR cfgDeviation_DB16) OR cfgDither_DB16) OR cfgPeriod_DB16) OR cfgPOC_DB16);
	status_b16: UINT;
	/// duty cycle 0..16#8000 
	dc_u16: UINT;
	///ADC digits, range from 0..25000
	digits_u16: UINT;
	/// set current [mA] 
	iSet_u16: UINT;
	/// actual current [mA] 
	iAct_u16: UINT;
	iActRaw_mA_u16: UINT;
	/// fault status 
	stDFC_SCB_u16: UINT;
	/// fault status 
	stDFC_SCG_u16: UINT;
	/// fault status 
	stDFC_OL_u16: UINT;
	/// fault status 
	stDFC_OT_u16: UINT;
	/// fault status 
	stDFC_OC_u16: UINT;
	/// fault status 
	stDFC_OR_u16: UINT;
	///Unintended switch ON of output
	unintendedSwitchONErr_l: BOOL;
	///locked by Inhibits
	lockedByINH_l: BOOL;
END_STRUCT
END_TYPE

// System API/SYS/STRUCTURE/bds_ResetInfo_ts
{attribute 'external_name' := 'cmp_rts_bds_ResetInfo_ts'}
TYPE bds_ResetInfo_ts :
STRUCT
	///User defined value, free for individual use, e.g. for Diagnostics.
	rbr_UserDefined_u32: UDINT;
	///Reset ID.
	rbr_Type_u16: UINT;
	///Reset group ID.
	rbr_Grp_u16: UINT;
	///Time stamp of current reset.
	rbr_TiStampCurr_u64: ULINT;
END_STRUCT
END_TYPE

// Diagnostics API/UDS/STRUCTURE/bds_uds_udsconfigparameter_ts
{attribute 'external_name' := 'cmp_rts_bds_uds_udsconfigparameter_ts'}
(*It is a structure which contains the details of UDS Node ID configuration, such as Node ID, Tester ID and Rx/Tx Identifiers for UDS message.*)
TYPE bds_uds_udsconfigparameter_ts :
STRUCT
	///Tester ID
	testerid_u8: USINT;
	///ECU Node ID
	nodeid_u8: USINT;
	///Rx and Tx Identifiers for the UDS message
	rxtxidentifiers_u16: UINT;
END_STRUCT
END_TYPE

// I/O API/IN legacy/STRUCTURE/bds_in_aiv_ts
{attribute 'external_name' := 'cmp_rts_bds_in_aiv_ts'}
TYPE bds_in_aiv_ts :
STRUCT
	///status flags for status_b16 
	///	
	///	initIn_DB16: USINT := 16#1;(*initialization after startup*)
	///	
	///	cfgAiv_DB16: USINT := 16#2;(*configured for AIV thresholds*)
	///	
	///	cfgAic_DB16: USINT := 16#4;(*configured for AIC thresholds*)
	///	
	///	cfgAid_DB16: USINT := 16#8;(*configured for AID thresholds*)
	///	
	///	cfgRi_DB16: USINT := 16#10;(*configured for RI thresholds*)
	///	
	///	cfgFreq_DB16: USINT := 16#20;(*configured for standard frequency sensor*)
	///	
	///	cfgFreqDSM_DB16: USINT := 16#40;(*configured for DSM frequency sensor*)
	///	
	///	lostSignalInfoDSM_DB16: USINT := 16#80;
	///	
	///	actShunt_DB16: UINT := 16#1000;(*shunt is activated for DSM sensor respective AIC*)
	///	
	///	lockReactShunt_DB16: UINT := 16#2000;(*locked shunt reactivation*)
	///	
	///	cfgInMask_DB16: UINT := (((((cfgFreqDSM_DB16 OR cfgFreq_DB16) OR cfgRi_DB16) OR cfgAid_DB16) OR cfgAic_DB16) OR cfgAiv_DB16);
	status_b16: UINT;
	///ADC digits, range from 0..25000 
	digits_u16: UINT;
	///voltage in [mV]
	u_mV_u16: UINT;
	///actual state 
	state_u8: USINT;
	///fault status
	stDFC_SCB_u16: UINT;
	///fault status
	stDFC_SCG_u16: UINT;
	///fault status
	stDFC_OR_u16: UINT;
END_STRUCT
END_TYPE

// Diagnostics API/UDS/UNION/bds_uds_udsconfigparameter_tu
{attribute 'external_name' := 'cmp_rts_bds_uds_udsconfigparameter_tu'}
(*It is a union which gives details about the Node ID parameters and CAN ID related data.*)
TYPE bds_uds_udsconfigparameter_tu :

UNION
	(*Structure which contains the UDS Node ID configuration parameters*)
	bds_uds_udsCfgPar_s: bds_uds_udsconfigparameter_ts;
	(*UDS CAN ID (Request)*)
	bds_uds_udsCanID_u32: UDINT;
END_UNION

END_TYPE

// I/O API/IN legacy/STRUCTURE/bds_in_sent_SDDataBox_ts
{attribute 'external_name' := 'cmp_rts_bds_in_sent_SDDataBox_ts'}
TYPE bds_in_sent_SDDataBox_ts :
STRUCT
	///This flag shows if the databox is initialised
	///   + FALSE: databox not initialised
	///   + TRUE : databox initialised	
	initialized_l: BOOL;
	///message identifier
	MsgID_u8: USINT;
	///start address of the buffer
	start_pas: POINTER TO bds_in_sent_slowData_ts;
	///Management of the buffer  
	Manage_s: bds_in_sent_BufManage_ts;
END_STRUCT
END_TYPE

// I/O API/IN legacy/STRUCTURE/bds_in_sent_slowData_ts
{attribute 'external_name' := 'cmp_rts_bds_in_sent_slowData_ts'}
TYPE bds_in_sent_slowData_ts :
STRUCT
	///Message ID  4 or 8 bit 
	MsgID_u8: USINT;
	///Data 12 or 16 bit
	Data_u16: UINT;
	///Status and Communication Nibble
	cfgBit_u8: USINT;
END_STRUCT
END_TYPE

// I/O API/IN legacy/STRUCTURE/bds_in_stPhase_ts
{attribute 'external_name' := 'cmp_rts_bds_in_stPhase_ts'}
TYPE bds_in_stPhase_ts :
STRUCT
	///frequency of the primary signal [dHz]
	frequency_u32: UDINT;
	///direction of rotation
	///   + 16#00 = left (ccw)
	///   + 16#01 = right (cw)
	direction_u8: USINT;
	///error status
	///   + 16#00 = error free or failure detection not possible
	///   + 16#01 = loss of primary signal or signal period is longer than status request 
	///   + 16#02 = loss of secondary signal 
	error_u8: USINT;
	///period primary signal [us]
	tiPeriodPrimSig_u32: UDINT;
	///period secondary signal [us]
	tiPeriodSecSig_u32: UDINT;
	///Time stamp [us] of rising edge of the primary signal
	tiPrimSig_u32: UDINT;
	///Time stamp [us] of rising edge of the secondary signal 
	tiSecSig_u32: UDINT;
	///phase shift of the signals [us]
	tiShift_u32: UDINT;
	///period counter - direction of counting depend on direction
	couPulse_s32: DINT;
	///state at function call time ("1" for high or "0" for low)
	stPrimSig_CurrSt_u8: USINT;
	///no update available (request within the same period)
	stPrimSig_samePer_u8: USINT;
	///period too long (timer overflow)
	stPrimSig_TimOvfl_u8: USINT;
	///measured period exceeds given maximum length 
	stPrimSig_MaxPerOvfl_u8: USINT;
	///state at function call time ("1" for high or "0" for low)
	stSecSig_CurrSt_u8: USINT;
	///no update available (request within the same period)
	stSecSig_samePer_u8: USINT;
	///period too long (timer overflow)
	stSecSig_TimOvfl_u8: USINT;
	///measured period exceeds given maximum length 
	stSecSig_MaxPerOvfl_u8: USINT;
	///Pointer of the start address of the period array primary signal 
	tiPeriodPrimSigExt_pcu32: POINTER TO UDINT;
	///Pointer of the start address of the pulse array primary signal 
	tiPulsePrimSigExt_pcu32: POINTER TO UDINT;
	///Pointer of the start address of the period array secondary signal 
	tiPeriodSecSigExt_pcu32: POINTER TO UDINT;
	///Pointer of the start address of the pulse array secondary signal 
	tiPulseSecSigExt_pcu32: POINTER TO UDINT;
END_STRUCT
END_TYPE

// System API/DSM/STRUCTURE/bds_dsm_j1939Lamp_ts
{attribute 'external_name' := 'cmp_rts_bds_dsm_j1939Lamp_ts'}
TYPE bds_dsm_j1939Lamp_ts :
STRUCT
	///lamp/flash status
	flash_state_u32: UDINT;
END_STRUCT
END_TYPE

// System API/DSM/STRUCTURE/bds_dsm_J1939_info_ts
{attribute 'external_name' := 'cmp_rts_bds_dsm_J1939_info_ts'}
TYPE bds_dsm_J1939_info_ts :
STRUCT
	///SPN for the DTC
	bds_SPN_u32: UDINT;
	///FMI for the DTC
	bds_FMI_u8: USINT;
	///Occurrence counter for the DTC
	bds_occur_count_u8: USINT;
	///Lamp State of DTC
	bds_lampState_u8: bds_dsm_j1939Lamp_ts;
END_STRUCT
END_TYPE

// System API/DSM/ENUM/bds_dsm_state_te
{attribute 'external_name' := 'cmp_rts_bds_dsm_state_te'}
TYPE bds_dsm_state_te :
(
	///Fault is Active.
	ACTIVE_ERRORS := 0,
	///Fault was Previously Active.
	PREVIOUSLY_ACTIVE_ERRORS
);
END_TYPE

// System API/SYS/STRUCTURE/bds_EcuInfo_ts
{attribute 'external_name' := 'cmp_rts_bds_EcuInfo_ts'}
TYPE bds_EcuInfo_ts :
STRUCT
	///Identification number of customer.
	IdNr_Custom_au8: ARRAY[1..19] OF USINT;
	///Identifier number BR SAP-ID_Number (Bosch Rexroth).
	IdNr_BR_au8: ARRAY[1..12] OF USINT;
	///Change revision AE (Automotive Electronics).
	ChangeRev_AE_au8: ARRAY[1..10] OF USINT;
	///Factory code.
	FactoryCode_au8: ARRAY[1..2] OF USINT;
	///Production date (YY-MM-DD).
	ProdDate_au8: ARRAY[1..3] OF USINT;
	///EEPROM version.
	Eeprom_Version_u8: USINT;
	///Calibration data.
	Calib_u8: USINT;
	///Hardware code.
	Hw_Typ_au8: ARRAY[1..2] OF USINT;
	///Serial number.
	SerialNr_au8: ARRAY[1..4] OF USINT;
	dummy_au8: ARRAY[1..2] OF USINT;
END_STRUCT
END_TYPE

// System API/DSM/STRUCTURE/bds_dsm_dfc_ts
{attribute 'external_name' := 'cmp_rts_bds_dsm_dfc_ts'}
TYPE bds_dsm_dfc_ts :
STRUCT
	/// REFERENCE number
	id: UINT := 12;
	/// assigned predebouncing mode
	debmode: UINT := 4;
END_STRUCT
END_TYPE

// System API/DSM/STRUCTURE/bds_dsm_dtcj1939_ts
{attribute 'external_name' := 'cmp_rts_bds_dsm_dtcj1939_ts'}
TYPE bds_dsm_dtcj1939_ts :
STRUCT
	///SPN value
	SPN_u32: UDINT;
	///FMI value
	FMI_u8: USINT;
	///lamp states
	lampState_u8: bds_dsm_j1939Lamp_ts;
END_STRUCT
END_TYPE

// System API/DSM/STRUCTURE/bds_dsm_fid_ts
{attribute 'external_name' := 'cmp_rts_bds_dsm_fid_ts'}
TYPE bds_dsm_fid_ts :
STRUCT
	///DFC reference ID
	id: UINT;
END_STRUCT
END_TYPE

// Communication API/ISOBUS/STRUCTURE/bds_isobus_appInst_ts
///Structure of a ISOBUS CA (controller application) instance.
{attribute 'external_name' := 'cmp_rts_bds_isobus_appInst_ts'}
TYPE bds_isobus_appInst_ts :
STRUCT
	/// user defined ISOBUS Receive data boxes info 
	rxDataboxInfo_s: bds_isobus_rxDataboxInfo_ts;
	/// user defined ISOBUS Transmit data boxes info
	txDataboxInfo_s: bds_isobus_txDataboxInfo_ts;
	//J1939-76 Producer databox
	prodDataboxInfo_s : bds_isobus_prodDataboxInfo_ts;
	//J1939-76 Consumer databox
	cnsrDataboxInfo_s : bds_isobus_cnsrDataboxInfo_ts;
	// Fixed transmission SDG data box handling
	prodSdgDataboxNum_u16 : UINT;
	// user defined CA address info table
    caAddrInfoTableRef_s  : bds_isobus_caAddrInfoTblRef_ts;
    // Callback pointer to indicate Addr Claim & Info table updates 
    addClaimInfoFunc_pf : POINTER TO UINT;  
	/// isobus tx bam control data
	txBamCtrl_s: bds_isobus_bamCtrl_ts;
	/// BAM message buffer for requestPGN answers
	txBamBuff_s: bds_isobus_txMsg_ts;
	/// rx tp control data for RTS/CTS transport layer
	rxTpCtrl_s: bds_isobus_rxTpCtrl_ts;
	/// tx tp control data for RTS/CTS transport layer
	txTpCtrl_s: bds_isobus_txTpCtrl_ts;
	/// rx ETP control data for RTS/CTS transport layer
	rxEtpCtrl_s: bds_isobus_rxEtpCtrl_ts;
	/// tx ETP control data for RTS/CTS transport layer
	txEtpCtrl_s: bds_isobus_txEtpCtrl_ts;
	/// function is called if DM3 msg received
	DM3func_pf: POINTER TO BOOL;
	/// function is called if DM11 msg received
	DM11func_pf: POINTER TO BOOL;
	/// pointer to ECU location string
	ecuLoc_pas8: POINTER TO SINT;
	/// pointer to ECU type string         
	ecuType_pas8: POINTER TO SINT;
	/// pointer to ECU manufacturer string
	ecuMan_pas8: POINTER TO SINT;
	/// pointer to application task name
	applTask_pas8: POINTER TO SINT;
	/// DM1/2 error data of own application
	err_s: bds_isobus_err_ts;
	/// internal isobus rx databoxes
	rxSysDatabox_as: ARRAY[1..5] OF bds_isobus_rxMsg_ts;
	/// internal isobus tx databoxes
	txSysDatabox_as: ARRAY[1..1] OF bds_isobus_txMsg_ts;
	/// data of rx databox for request PGN msg
	rxDataRequPgn_au8: ARRAY[1..8] OF USINT;
	/// data of rx databox for address claim msg
	rxDataAddrClm_au8: ARRAY[1..8] OF USINT;
	/// data of rx databox for commanded msg
	rxDataCmdAddr_au8: ARRAY[1..9] OF USINT;
	/// data of rx databox for name management msg
	rxDataNameNmt_au8: ARRAY[1..8] OF USINT;
	/// data of rx databox for DM13 msg
	rxDataDm13_au8: ARRAY[1..8] OF USINT;
	/// tx buffer for RequPgn msg
	txDataRequPgn_au8: ARRAY[1..300] OF USINT;
	/// buffer for DM1 tx databox
	dm1BuffDat_au8: ARRAY[1..130] OF USINT;
	/// buffer for DM2 tx databox
	dm2BuffDat_au8: ARRAY[1..130] OF USINT;
	/// controller application name
	caName_u: bds_isobus_caName_tu;
	/// controller application pending name
	caPendName_u: bds_isobus_caName_tu;
	/// global status of controller application
	caStatus_u16: UINT;
	/// timer [ms] for address claiming supervision
	addrClaimTimer_u16: UINT;
	/// Periodic databox array index for continuing transmission in next cycle
	taskNxtPeriodicTxIdx_u16: UINT;
	/// own CA (source) address
	ownAddr_u8: USINT;
	/// can channel used by CA
	canChannel_u8: USINT;
	/// source address of last name management request
	nameMngSourceAddr_u8: USINT;
	/// port (0..11) to be evaluated from DM13 message
	usedDm13Port_u8: USINT;
	/// TRUE, if add. DM1 may be sent wihtin 1s periode
	sendDm1Allowed_l: BOOL;
	///TRUE -> handle DM1/DM2 lamp state according J1939
	dmLampStateJ1939_l: BOOL;
	aperiodicDataboxNum_s: bds_isobus_aperiodicDataboxNum_ts; // Aperiodic Databox Handling
    periodicDataboxNum_s: bds_isobus_periodicDataboxNum_ts;  // Periodic Databox Handling

END_STRUCT
END_TYPE

// Communication API/ISOBUS/STRUCTURE/bds_isobus_bamCtrl_ts
///Struct for isobus BAM transport control
{attribute 'external_name' := 'cmp_rts_bds_isobus_bamCtrl_ts'}
TYPE bds_isobus_bamCtrl_ts :
STRUCT
	///nbr already sent data bytes
	lenTx_u16: UINT;
	///timer for TX BAM control
	timer_u16: UINT;
	///status of TX BAM protocol handler
	state_u8: USINT;
	///ptr to message buffer, which is currently sended via BAM
	txMsg_ps: POINTER TO bds_isobus_txMsg_ts;
END_STRUCT
END_TYPE

// Communication API/ISOBUS/STRUCTURE/bds_isobus_caName_ts
///Structure of CA name
{attribute 'external_name' := 'cmp_rts_bds_isobus_caName_ts'}
TYPE bds_isobus_caName_ts :
STRUCT
	caName_u32: UDINT;
END_STRUCT
END_TYPE

// Communication API/ISOBUS/UNION/bds_isobus_caName_tu
{attribute 'external_name' := 'cmp_rts_bds_isobus_caName_tu'}
TYPE bds_isobus_caName_tu :

UNION
	name_au8: ARRAY[1..8] OF USINT;
	name_s: bds_isobus_caName_ts;
	nm_s: bds_isobus_nm_ts;
END_UNION

END_TYPE

// Communication API/ISOBUS/STRUCTURE/bds_isobus_canID_ts
{attribute 'external_name' := 'cmp_rts_bds_isobus_canID_ts'}
TYPE bds_isobus_canID_ts :
STRUCT
	bitFormat_u32: UDINT;
END_STRUCT
END_TYPE

// Communication API/ISOBUS/UNION/bds_isobus_canID_tu
{attribute 'external_name' := 'cmp_rts_bds_isobus_canID_tu'}
TYPE bds_isobus_canID_tu :
UNION
	canID_s : bds_isobus_canID_ts;
	canID_u32 : UDINT;
END_UNION
END_TYPE

// I/O API/IN legacy/STRUCTURE/bds_in_ri_ts
{attribute 'external_name' := 'cmp_rts_bds_in_ri_ts'}
TYPE bds_in_ri_ts :
STRUCT
	///status flags for status_b16 
	///	
	///	initIn_DB16: USINT := 16#1;(*initialization after startup*)
	///	
	///	cfgAiv_DB16: USINT := 16#2;(*configured for AIV thresholds*)
	///	
	///	cfgAic_DB16: USINT := 16#4;(*configured for AIC thresholds*)
	///	
	///	cfgAid_DB16: USINT := 16#8;(*configured for AID thresholds*)
	///	
	///	cfgRi_DB16: USINT := 16#10;(*configured for RI thresholds*)
	///	
	///	cfgFreq_DB16: USINT := 16#20;(*configured for standard frequency sensor*)
	///	
	///	cfgFreqDSM_DB16: USINT := 16#40;(*configured for DSM frequency sensor*)
	///	
	///	lostSignalInfoDSM_DB16: USINT := 16#80;
	///	
	///	actShunt_DB16: UINT := 16#1000;(*shunt is activated for DSM sensor respective AIC*)
	///	
	///	lockReactShunt_DB16: UINT := 16#2000;(*locked shunt reactivation*)
	///	
	///	cfgInMask_DB16: UINT := (((((cfgFreqDSM_DB16 OR cfgFreq_DB16) OR cfgRi_DB16) OR cfgAid_DB16) OR cfgAic_DB16) OR cfgAiv_DB16);
	status_b16: UINT;
	///ADC digits, range from 0..25000
	digits_u16: UINT;
	///voltage in [mV]
	u_mV_u16: UINT;
	///resistance in [R]
	ohm_r_u32: UDINT;
	///fault status
	stDFC_SCB_u16: UINT;
	///fault status
	stDFC_SCG_u16: UINT;
	///temperature [°C]
	tCelsius_s16: INT;
END_STRUCT
END_TYPE

// I/O API/IN legacy/STRUCTURE/bds_in_sent_BufManage_ts
{attribute 'external_name' := 'cmp_rts_bds_in_sent_BufManage_ts'}
TYPE bds_in_sent_BufManage_ts :
STRUCT
	length_u16: UINT;
	idx_in_u16: UINT;
	idx_out_u16: UINT;
	BufEmpty_l: BOOL;
	BufOvfl_l: BOOL;
END_STRUCT
END_TYPE

// I/O API/IN legacy/STRUCTURE/bds_in_sent_copyFDBuf_ts
{attribute 'external_name' := 'cmp_rts_bds_in_sent_copyFDBuf_ts'}
TYPE bds_in_sent_copyFDBuf_ts :
STRUCT
	/// length of copy buffer
	lengthCopyBuf_u8: USINT;
	/// pointer to copy buffer 
	start_pas: POINTER TO bds_in_sent_decodedFD_ts;
	///actual length of buffer
	length_u8: USINT;
	///This flag shows if the buffer is completely filled
	///   + FALSE: until now the buffer is not full
	///   + TRUE : buffer is full
	full_l: BOOL;
END_STRUCT
END_TYPE

// I/O API/IN legacy/STRUCTURE/bds_in_sent_databoxinfo_ts
{attribute 'external_name' := 'cmp_rts_bds_in_sent_databoxinfo_ts'}
TYPE bds_in_sent_databoxinfo_ts :
STRUCT
	num_u8: USINT;
	mem_pas: POINTER TO bds_in_sent_SDDataBox_ts;
END_STRUCT
END_TYPE

// Communication API/ISOBUS/STRUCTURE/bds_isobus_dtcList_ts
///Structure of received and converted DM1/2 failure lists
{attribute 'external_name' := 'cmp_rts_bds_isobus_dtcList_ts'}
TYPE bds_isobus_dtcList_ts :
STRUCT
	///lamp status
	lamp_s: bds_isobus_lamp_ts;
	///DTC list
	dtc_as: ARRAY[1..20] OF bds_isobus_dtc_ts;
END_STRUCT
END_TYPE

// I/O API/IN legacy/STRUCTURE/bds_in_sent_decodedFD_ts
{attribute 'external_name' := 'cmp_rts_bds_in_sent_decodedFD_ts'}
TYPE bds_in_sent_decodedFD_ts :
STRUCT
	/// channel 1 data 
	chnl1Val_u16: UINT;
	///optional channel 2 data 
	chnl2Val_u16: UINT;
	///optional counter 
	counter_u8: USINT;
	///optional inverted channel 1 MSN 
	invMSN_u8: USINT;
	///Message / Status nibble 
	msgStat_u8: USINT;
END_STRUCT
END_TYPE

// Communication API/ISOBUS/STRUCTURE/bds_isobus_dtc_ts
///Structure of one DTC
{attribute 'external_name' := 'cmp_rts_bds_isobus_dtc_ts'}
TYPE bds_isobus_dtc_ts :
STRUCT
	///suspect parameter number
	spn_u32: UDINT;
	///failure mode indicator
	fmi_u8: USINT;
	///occurrence counter
	occ_u8: USINT;
END_STRUCT
END_TYPE

// Communication API/ISOBUS/STRUCTURE/bds_isobus_err_ts
///Structure of all data for one error handler instance for DM1 and DM2 failures
{attribute 'external_name' := 'cmp_rts_bds_isobus_err_ts'}
TYPE bds_isobus_err_ts :
STRUCT
	///TX box nbr for sending the DM1 failures
	txBoxDM1_u16: UINT;
	///TX box nbr for sending the DM2 failures
	txBoxDM2_u16: UINT;
END_STRUCT
END_TYPE

// Communication API/ISOBUS/STRUCTURE/bds_isobus_rxDataboxInfo_ts
///Structure of isobus rx data box info for API
{attribute 'external_name' := 'cmp_rts_bds_isobus_rxDataboxInfo_ts'}
TYPE bds_isobus_rxDataboxInfo_ts :
STRUCT
	///pointer to the buffer for data boxes
	mem_pas: POINTER TO bds_isobus_rxMsg_ts;
	///number of data boxes
	num_u16: UINT;
END_STRUCT
END_TYPE

// Communication API/ISOBUS/STRUCTURE/bds_isobus_rxEtpCtrl_ts
///Structure with required data for receiving rx databox via ETP handler
{attribute 'external_name' := 'cmp_rts_bds_isobus_rxEtpCtrl_ts'}
TYPE bds_isobus_rxEtpCtrl_ts :
STRUCT
	///response or transmit CANid
	canID_u: bds_isobus_canID_tu;
	///PGN to be handled
	PGN_u32: UDINT;
	///pointer to rx databox, currently handled by mtp handler
	rxMsgPtr_ps: POINTER TO bds_isobus_rxMsg_ts;
	///nbr of already handled data bytes of succ. completed packages
	doneDataCnt_u32: UDINT;
	///first message (=offset) nbr of the package to be handled
	packageStart_u32: UDINT;
	///last message number = total nbr of messages
	lastPackage_u32: UDINT;
	///time counter [ms] for timeout supervision
	timer_u16: UINT;
	///actual message sequence number to be received
	packageNumber_u8: USINT;
	///nbr of single msgs per burst which fit into buffer
	packageCount_u8: USINT;
	///max. nbr of messages to be handled per burst (for CTS msg)
	maxPackage_u8: USINT;
	///status of state machine
	state_u8: USINT;
	///retry flag for requesting the same package via CTS
	retryCtsFlag_l: BOOL;
END_STRUCT
END_TYPE

// Communication API/ISOBUS/STRUCTURE/bds_isobus_rxMsg_ts
///Structure of a isobus rx databox message definition within the array of defined rx messages
{attribute 'external_name' := 'cmp_rts_bds_isobus_rxMsg_ts'}
TYPE bds_isobus_rxMsg_ts :
STRUCT
	///pointer to data array with length=lenMax_u32
	data_pau8: POINTER TO USINT;
	///function is called if msg received completely
	func_pf: POINTER TO BOOL;
	///can identity of msg to be received
	canID_u: bds_isobus_canID_tu;
	///expected total length of actual received msg to be receievd
	lenAct_u32: UDINT;
	///length of already received msg part
	lenRx_u32: UDINT;
	///max length of the receive buffer
	lenMax_u32: UDINT;
	///timeout (ms) for supervision of cyclic msg
	timeout_u16: UINT;
	///start timeout (ms) for supervision of first msg
	startTimeout_u16: UINT;
	///actual time counter for timeout supervision
	counter_u16: UINT;
	///msg status, e.g. valid, invalid, timeout
	status_u16: UINT;
	///action (e.g. data conversion) to be done after reception
	action_u16: UINT;
	///= true, if it is an stack internal rx databox
	internalBox_l: BOOL;
END_STRUCT
END_TYPE

// Communication API/ISOBUS/STRUCTURE/bds_isobus_rxTpCtrl_ts
///Structure with required data for receiving rx databox via mtp handler
{attribute 'external_name' := 'cmp_rts_bds_isobus_rxTpCtrl_ts'}
TYPE bds_isobus_rxTpCtrl_ts :
STRUCT
	///Response or transmit CANid
	canID_u: bds_isobus_canID_tu;
	///PGN to be handled
	PGN_u32: UDINT;
	///Pointer to rx databox, currently handled by mtp handler
	rxMsgPtr_ps: POINTER TO bds_isobus_rxMsg_ts;
	///Nbr of already handled data bytes OF succ. completed packages
	doneDataCnt_u16: UINT;
	///Time counter [ms] for timeout supervision
	timer_u16: UINT;
	///Nbr of single msgs (packets) per package which fit into buff.
	packageCount_u8: USINT;
	///First message (packet) nbr of the package to be handled
	packageStart_u8: USINT;
	///Actual message sequence (packet) number
	packageNumber_u8: USINT;
	///Last message (packet) number
	lastPackage_u8: USINT;
	///Max. nbr of messages to be handled per packet (for CTS msg)
	maxPackage_u8: USINT;
	///Status of state machine
	state_u8: USINT;
	///Retry flag for requesting the same package via CTS
	retryCtsFlag_l: BOOL;
END_STRUCT
END_TYPE

// Communication API/ISOBUS/STRUCTURE/bds_isobus_txDataboxInfo_ts
///Structure of isobus tx data box info for API.
{attribute 'external_name' := 'cmp_rts_bds_isobus_txDataboxInfo_ts'}
TYPE bds_isobus_txDataboxInfo_ts :
STRUCT
	/// Pointer to the buffer for data boxes
	mem_pas: POINTER TO bds_isobus_txMsg_ts;
	/// Number of data boxes
	num_u16: UINT;
END_STRUCT
END_TYPE

// Communication API/ISOBUS/STRUCTURE/bds_isobus_txEtpCtrl_ts
///Structure with required data for transmitting tx databox via ETP handler
{attribute 'external_name' := 'cmp_rts_bds_isobus_txEtpCtrl_ts'}
TYPE bds_isobus_txEtpCtrl_ts :
STRUCT
	///Response or transmit CANid
	canID_u: bds_isobus_canID_tu;
	///PGN to be handled
	PGN_u32: UDINT;
	/// Pointer to tx databox, currently handled by mtp handler
	txMsgPtr_ps: POINTER TO bds_isobus_txMsg_ts;
	/// Total number of data bytes
	msgDlc_u32: UDINT;
	/// Nbr of already handled data bytes
	doneDataCnt_u32: UDINT;
	/// First message (=offset) nbr of the package to be handled
	packageStart_u32: UDINT;
	/// Last message number = total nbr of messages
	lastPackage_u32: UDINT;
	/// Time counter [ms] for timeout supervision
	timer_u16: UINT;
	/// Actual message sequence number
	packageNumber_u8: USINT;
	/// Nbr of msgs for next burst which must fit into buffer
	packageCount_u8: USINT;
	/// Max. nbr of messages to be handled per burst (for CTS msg)
	maxPackage_u8: USINT;
	/// Status of state machine
	state_u8: USINT;
END_STRUCT
END_TYPE

// Communication API/ISOBUS/STRUCTURE/bds_isobus_txMsg_ts
///Structure of a isobus tx databox message definition within the array of defined tx messages
{attribute 'external_name' := 'cmp_rts_bds_isobus_txMsg_ts'}
TYPE bds_isobus_txMsg_ts :
STRUCT
	/// Pointer to data array with length=lenMax_u32
	data_pau8: POINTER TO USINT;
	/// Function is called before msg is to be sent
	func_pf: POINTER TO UDINT;
	/// CAN identity of msg to be sent
	canID_u: bds_isobus_canID_tu;
	/// Max length (buffer size) of msg to be sent
	lenMax_u32: UDINT;
	/// Actual length of msg to be sent
	lenAct_u32: UDINT;
	/// Cycle time for sending this msg
	cycle_u16: UINT;
	/// Cycle time for sending this msg
	counter_u16: UINT;
	/// Msg status, e.g. valid, invalid
	status_u16: UINT;
	aperiodicdatabox_u16: UINT;
	periodicdatabox_u16: UINT;
END_STRUCT
END_TYPE

// Communication API/ISOBUS/STRUCTURE/bds_isobus_txTpCtrl_ts
{attribute 'external_name' := 'cmp_rts_bds_isobus_txTpCtrl_ts'}
TYPE bds_isobus_txTpCtrl_ts :
STRUCT
	/// Response or transmit CANid
	canID_u: bds_isobus_canID_tu;
	/// PGN to be handled
	PGN_u32: UDINT;
	/// Pointer to tx databox, currently handled by mtp handler
	txMsgPtr_ps: POINTER TO bds_isobus_txMsg_ts;
	/// Total number of data bytes
	msgDlc_u16: UINT;
	/// Nbr of already handled data bytes
	doneDataCnt_u16: UINT;
	/// Time counter [ms] for timeout supervision
	timer_u16: UINT;
	/// Nbr of single msgs (packets) per package which fit into buff.
	packageCount_u8: USINT;
	/// First message (packet) nbr of the package to be handled
	packageStart_u8: USINT;
	/// Actual message sequence number to be sent
	packageNumber_u8: USINT;
	/// Last message (packet) number
	lastPackage_u8: USINT;
	/// Status of state machine
	state_u8: USINT;
END_STRUCT
END_TYPE

// Communication API/ISOBUS/STRUCTURE/bds_isobus_lamp_ts
///Structure of one lamp status
{attribute 'external_name' := 'cmp_rts_bds_isobus_lamp_ts'}
TYPE bds_isobus_lamp_ts :
STRUCT
	///lamp status
	lampState_u8: USINT;
	///lamp flash
	lampFlash_u8: USINT;
END_STRUCT
END_TYPE

// Communication API/ISOBUS/STRUCTURE/bds_isobus_nm_ts
///Structure for name management services
{attribute 'external_name' := 'cmp_rts_bds_isobus_nm_ts'}
TYPE bds_isobus_nm_ts :
STRUCT
	nameManagement_u32: UDINT;
END_STRUCT
END_TYPE

// I/O API/OUT/STRUCTURE/bds_out_aov_ts
{attribute 'external_name' := 'cmp_rts_bds_out_aov_ts'}
TYPE bds_out_aov_ts :
STRUCT
	///status flags for status_b16 
	///	initOut_DB16: USINT := 16#1;(*initialization after startup*)
	///	
	///	cfgPOC_DB16: USINT := 16#2;(*configuration of closed loop control*)
	///	
	///	cfgPeriod_DB16: USINT := 16#4;(*configuration of period*)
	///	
	///	cfgDither_DB16: USINT := 16#8;(*configuration of dither*)
	///	
	///	cfgDeviation_DB16: USINT := 16#10;(*configuration of deviation*)
	///	
	///	cfgPI_DB16: USINT := 16#20;(*configuration of KpKi*)
	///	
	///	lockedSCB_DB16: USINT := 16#40;(*locked by SCB...necessary for AOV*)
	///	
	///	lockedSCG_DB16: USINT := 16#80;(*locked by SCG...necessary for AOV*)
	///	
	///	lockedOC_DB16: UINT := 16#100;(*locked by OC*)
	///	
	///	locked_DB16: UINT := 16#200;(*locked by Error Handler*)
	///	
	///	lockedMO_DB16: UINT := 16#400;(*locked by Monitoring Module (MO) Error*)
	///	
	///	lockCouTiReact_DB16: UINT := 16#800;(*locked reactivation timer reload after a hot short circuit*)
	///	
	///	tiReactNotElapsed_DB16: UINT := 16#1000;(*time for reactivation after a hot short circuit not elapsed*)
	///	
	///	linked_DB16: UINT := 16#2000;(*linked at least with one other safout output*)
	///	
	///	tlsPlsDis_DB16: UINT:=16#4000;(*Test pulses disable*)
	///	
	///	disabled_DB16: UINT := 16#8000;(*output is disabled (avoid open load faults of unused outputs)*)
	///	
	///	cfgOutMask_DB16: UINT := ((((cfgPI_DB16 OR cfgDeviation_DB16) OR cfgDither_DB16) OR cfgPeriod_DB16) OR cfgPOC_DB16);
	status_b16: UINT;
	///duty cycle 0..1000 [0,1%]
	dc_u16: UINT;
	///ADC digits, range from 0..25000
	digits_u16: UINT;
	///setpoint voltage [mV]
	uSet_u16: UINT;
	///actual voltage [mV]
	uAct_u16: UINT;
	///fault status
	stDFC_SCB_u16: UINT;
	///fault status
	stDFC_SCG_u16: UINT;
	///fault status
	stDFC_OR_u16: UINT;
END_STRUCT
END_TYPE

// I/O API/IN legacy/STRUCTURE/bds_in_sent_FDBufInfo_ts
{attribute 'external_name' := 'cmp_rts_bds_in_sent_FDBufInfo_ts'}
TYPE bds_in_sent_FDBufInfo_ts :
STRUCT
	start_pas: POINTER TO bds_in_sent_decodedFD_ts;
	Manage_s: bds_in_sent_BufManage_ts;
END_STRUCT
END_TYPE

// I/O API/OUT/ENUM/bds_load_characteristic_te
{attribute 'external_name' := 'cmp_rts_bds_load_characteristic_te'}
TYPE bds_load_characteristic_te :
(
	INDUCTIVE_LOAD := 0,
	CAPACITIVE_LOAD := 1
)USINT;
END_TYPE

// I/O API/IN legacy/STRUCTURE/bds_in_phase_ts
{attribute 'external_name' := 'cmp_rts_bds_in_phase_ts'}
TYPE bds_in_phase_ts :
STRUCT
	///frequency of the primary signal [dHz]
	frequency_u32: UDINT;
	///direction of rotation 
	///   + 16#00 = left (ccw)
	///   + 16#01 = right (cw) 
	direction_u8: USINT;
END_STRUCT
END_TYPE

// System API/SYS/ENUM/bds_sysCmn_status_te
{attribute 'external_name' := 'cmp_rts_bds_sysCmn_status_te'}
(*Enumeration listing the different return values possible for Post Build Selectable feature.*)
TYPE bds_sysCmn_status_te :
(
	(*Success : API executed without error*)
    bds_sysCmn_ok_E:= 0,
	(*Input variant is invalid*)
    bds_sysCmn_invalidVrnt_E,
	(*Variant is already configured, re-configuration is requested.*)
    bds_sysCmn_vrntReCfg_E
);
END_TYPE

// System API/SYS/STRUCTURE/bds_sysPb_retValCfgVrnt_ts
{attribute 'external_name' := 'cmp_rts_bds_sysPb_retValCfgVrnt_ts'}
(*Structure listing the return value for API related to |bds_sysPb_cfgVariant|.*)
TYPE bds_sysPb_retValCfgVrnt_ts :
STRUCT
	(*All possible return values are listed as Enumeration.*)
	status_e: bds_sysCmn_status_te;
END_STRUCT
END_TYPE

// System API/SYS/STRUCTURE/bds_sysPb_vrntParam_ts
{attribute 'external_name' := 'cmp_rts_bds_sysPb_vrntParam_ts'}
(*Structure which contains all the variants which shall be configured through easyConfig.*)
TYPE bds_sysPb_vrntParam_ts :
STRUCT
	(*This is the enum which contains the variants list.*)
	returnVrnt_te: usint;
END_STRUCT
END_TYPE

// System API/SYS/STRUCTURE/bds_sysPb_retValGetVrnt_ts
{attribute 'external_name' := 'cmp_rts_bds_sysPb_retValGetVrnt_ts'}
(*Structure listing the variants, related to |bds_sysPb_getVariant|.*)
TYPE bds_sysPb_retValGetVrnt_ts :
STRUCT
	(*List of variants configured in the project.Import bds_rts_ec.xml to use the enum bds_sysPb_vrnt_te.*)
	returnVrnt_te: usint;
END_STRUCT
END_TYPE

// I/O API/SENT/STRUCTURE/bds_sent_chSt_tb
(*Bit field type definition for the SENT module with status information of SENT functionality.
These bits will be set or reset based on the SENT Fast or Slow message received and SENT driver status.*)
{attribute 'external_name' := 'cmp_rts_bds_sent_chSt_tb'}
TYPE bds_sent_chSt_tb :
STRUCT
	initDrvr_b1: BIT;
	runngDrvr_b1: BIT;
	oneFrmRxd_b1: BIT;
	newFrmRxd_b1: BIT;
	oneSlowFrmRxd_b1: BIT;
	newSlowFrmRxd_b1: BIT;
	lineLo_b1: BIT;
	lineHi_b1: BIT;
	noDataRxd_b1: BIT;
	noEdgeRxd_b1: BIT;
	noiseDetd_b1: BIT;
	debd_b1: BIT;
	crcErr_b1: BIT;
	nibbleRngErr_b1: BIT;
	missNibble_b1: BIT;
	ovfNibble_b1: BIT;
	msgLost_b1: BIT;
	slowChCrcErr_b1: BIT;
	slowChMissFrm_b1: BIT;
	slowChNoDataRxd_b1: BIT;
	calibrationPlsOutOfRng_b1: BIT;
	calibrationPlsRepDe_b1: BIT;
	resd0_b1: BIT;
	breakPlsOutOfRng_b1: BIT;
	fastDataCntrErr_b1: BIT;
	fastDataInvtNibbleErr_b1: BIT;
	msgLostHwOverrun_b1: BIT;
	resd1_b1: BIT;
	resd2_b1: BIT;
	resd3_b1: BIT;
	resd4_b1: BIT;
	resd5_b1: BIT;
END_STRUCT
END_TYPE

// I/O API/SENT/ENUM/bds_sentCmn_status_te
(*Enumeration encoding the result status of the SENT API functions.*)
{attribute 'external_name' := 'cmp_rts_bds_sentCmn_status_te'}
TYPE bds_sentCmn_status_te :
(
	(*Call successful and signal can be used *)
	bds_sentCmn_ok_E := 0,
	(*Signal out of range (e.g., maximum period exceeded)*)
    bds_sentCmn_outOfRng_E,
	(*No measurement available due to external conditions (e.g., SENT channel is not running)*)
    bds_sentCmn_errExt_E,
	(*Not available (e.g., no Fast or Slow SENT message received, called to early in initialization phase, system in a mode it cannot measure etc.)*)
    bds_sentCmn_notAvl_E,
	(*Not available due to an internal error (e.g., SENT broken)*)
    bds_sentCmn_errInt_E,
	(*API call invalid, configuration invalid for the requested signal, etc.*)
    bds_sentCmn_invldCfg_E,
	(*API call invalid, incorrect parameters.*)
    bds_sentCmn_invldPrm_E
)USINT;
END_TYPE

// I/O API/SENT/STRUCTURE/bds_sent_rxFastData_ts
(*Data structure for latest received SENT Fast Data message of the API function |bds_sent_getFastData|.*)
{attribute 'external_name' := 'cmp_rts_bds_sent_rxFastData_ts'}
TYPE bds_sent_rxFastData_ts :
STRUCT
	(*SENT driver status information in bit format*)
	chSt_b: bds_sent_chSt_tb ;
	(*Array of all SENT received raw single Fast Data nibbles*)
	rxFastData_au8: ARRAY[1..8] OF USINT;
	(*Function call status return value*)
	status_e: bds_sentCmn_status_te;
END_STRUCT
END_TYPE

// I/O API/SENT/STRUCTURE/bds_sent_rxSlowData_ts
(*Data structure for latest received SENT Slow Data message of the API function |bds_sent_getSlowData|.*)
{attribute 'external_name' := 'cmp_rts_bds_sent_rxSlowData_ts'}
TYPE bds_sent_rxSlowData_ts :
STRUCT
	(*SENT driver status information in bit format*)
	chSt_b: bds_sent_chSt_tb;
	(*Slow Data 12 or 16 bit*)
	rxSlowData_u32: UDINT;
	(*Message ID 4 or 16 bit*)
	msgId_u8: USINT;
	(*Configuration bit*)
	cfgBit_u8: USINT;
	(*Function call status return value*)
	status_e:bds_sentCmn_status_te;
END_STRUCT
END_TYPE

// I/O API/SENT/STRUCTURE/bds_sent_getSlowDataBufd_ts
(*Data structure for a number of received SENT Slow Data frame samples of the API function |bds_sent_getSlowDataBufd|.*)
{attribute 'external_name' := 'cmp_rts_bds_sent_getSlowDataBufd_ts'}
TYPE bds_sent_getSlowDataBufd_ts :
STRUCT
	(*SENT driver status information in bit format*)
	chSt_b: bds_sent_chSt_tb;
	(*Number of received Slow Data samples since last function call, if Slow Data Buffer overflow the buffer size defined in easyConfig will be set.*)
	cntNewSample_u8: USINT;
	(*Function call status return value*)
	status_e:bds_sentCmn_status_te;
END_STRUCT
END_TYPE

// I/O API/SENT/STRUCTURE/bds_sent_getFastDataBufd_ts
(*Data structure for a number of received SENT Fast Data frame samples of the API function |bds_sent_getFastDataBufd|.*)
{attribute 'external_name' := 'cmp_rts_bds_sent_getFastDataBufd_ts'}
TYPE bds_sent_getFastDataBufd_ts :
STRUCT
	(*SENT driver status information in bit format*)
	chSt_b: bds_sent_chSt_tb;
	(*Number of received Fast Data samples since last function call, if Fast Data Buffer overflow the buffer size defined in easyConfig will be set*)
	cntNewSample_u8: USINT;
	(*Function call status return value*)
	status_e:bds_sentCmn_status_te;
END_STRUCT
END_TYPE

// I/O API/SENT/STRUCTURE/bds_sent_fastDataMsg_ts
(*Data structure type definition for received message Fast Data nibbles of one received sample.*)
{attribute 'external_name' := 'cmp_rts_bds_sent_fastDataMsg_ts'}
TYPE bds_sent_fastDataMsg_ts :
STRUCT
	(*Array for Fast Data Nibbles of one received sample*)
	rxFastData_au8: ARRAY[1..8] OF USINT;
END_STRUCT
END_TYPE

// I/O API/SENT/STRUCTURE/bds_sent_fastDataBuf_ts
(*Data structure type definition for received Fast Data Buffered messages of the API function bds_sent_getFastDataBufd.*)
{attribute 'external_name' := 'cmp_rts_bds_sent_fastDataBuf_ts'}
TYPE bds_sent_fastDataBuf_ts :
STRUCT
	(*Array for Fast Data Buffered values*)
	fastDataBufd_as: ARRAY[1..20] OF bds_sent_fastDataMsg_ts;
END_STRUCT
END_TYPE

// I/O API/SENT/STRUCTURE/bds_sent_slowDataMsg_ts
(*Data structure type definition for received message Slow Data of one received sample.*)
{attribute 'external_name' := 'cmp_rts_bds_sent_slowDataMsg_ts'}
TYPE bds_sent_slowDataMsg_ts :
STRUCT
	(*Received Slow Data 12 or 16 bit*)
	rxSlowData_u32: UDINT;
	(*Slow Data Message Identifier 4 or 8 bit*)
	msgId_u8: USINT;
	(*Slow Data status and communication nibble*)
	cfgBit_u8: USINT;
END_STRUCT
END_TYPE

// I/O API/SENT/STRUCTURE/bds_sent_slowDataBuf_ts
(*Data structure type definition for received Slow Data Buffered messages of the API function |bds_sent_getSlowDataBufd|.*)
{attribute 'external_name' := 'cmp_rts_bds_sent_slowDataBuf_ts'}
TYPE bds_sent_slowDataBuf_ts :
STRUCT
	(*Array type definition of Slow Data Messages*)
	slowDataBufd_as: ARRAY[1..20] OF bds_sent_slowDataMsg_ts;
END_STRUCT
END_TYPE

// I/O API/IN/STRUCTURE/bds_inI_measmt_ts
(*Data structure for one current measurement value of the API function |bds_inI_get|.*)
{attribute 'external_name' := 'cmp_rts_bds_inI_measmt_ts'}
TYPE bds_inI_measmt_ts :
STRUCT
	(*Measured current in micro Ampere*)
	i_uA_u16: UINT;
	(*Shunt state of the input current measurement signal*)
	stShunt_e: bds_inI_stShunt_te;
	(*Status of the measurement*)
	status_e: bds_inCmn_status_te;	
END_STRUCT
END_TYPE

// I/O API/IN/STRUCTURE/bds_inDig_measmt_ts
(*Data structure for one digital measurement value of the API function |bds_inDig_get|.*)
{attribute 'external_name' := 'cmp_rts_bds_inDig_measmt_ts'}
TYPE bds_inDig_measmt_ts :
STRUCT
	(*Digital state of input is high (0 = OFF, 1 = ON)*)
	stHigh_l: BOOL;
	(*Status of the measurement*)
	status_e: bds_inCmn_status_te;	
END_STRUCT
END_TYPE

// I/O API/IN/STRUCTURE/bds_inCmn_pullParam_ts
(*Data structure for input parameters for the API function |bds_inU_cfgPull|, |bds_inDig_cfgPull| and |bds_inI_cfgPull|.*)
{attribute 'external_name' := 'cmp_rts_bds_inCmn_pullParam_ts'}
TYPE bds_inCmn_pullParam_ts :
STRUCT
	(*Pull type*)
	pullType_e: bds_inCmn_pullType_te;
	(*Pull current strength *)
	iPull_e: bds_inCmn_iPull_te;
END_STRUCT
END_TYPE

// I/O API/IN/STRUCTURE/bds_inI_cfgPull_ts
(*Return structure for the API function |bds_inI_cfgPull|.*)
{attribute 'external_name' := 'cmp_rts_bds_inI_cfgPull_ts'}
TYPE bds_inI_cfgPull_ts :
STRUCT
	(*Status of the API call*)
	status_e: bds_inCmn_status_te;	
END_STRUCT
END_TYPE

// I/O API/IN/STRUCTURE/bds_inI_shunt_ts
(*Return structure of the API function |bds_inI_ctrlShunt|.*)
{attribute 'external_name' := 'cmp_rts_bds_inI_shunt_ts'}
TYPE bds_inI_shunt_ts :
STRUCT
	(*Status of function call to control the shunt*)
	status_e: bds_inCmn_status_te;	
END_STRUCT
END_TYPE

// I/O API/IN/STRUCTURE/bds_inDig_cfgPull_ts
(*Return structure for the API function |bds_inDig_cfgPull|.*)
{attribute 'external_name' := 'cmp_rts_bds_inDig_cfgPull_ts'}
TYPE bds_inDig_cfgPull_ts :
STRUCT
	(*Status of the API call*)
	status_e: bds_inCmn_status_te;	
END_STRUCT
END_TYPE

// I/O API/IN/ENUM/bds_inCmn_status_te
(*Enumeration encoding the result status of the input API functions.*)
{attribute 'external_name' := 'cmp_rts_bds_inCmn_status_te'}
TYPE bds_inCmn_status_te :
(
	(*Call successful and signal can be used*)
	bds_inCmn_ok_E := 0,
	(*Signal out of range (e.g., maximum period exceeded)*)
    bds_inCmn_outOfRng_E,
	(*No measurement available due to external conditions (e.g., UBat too low for ADC measurement)*)
    bds_inCmn_errExt_E,
	(*Not available (e.g., busy, called to early in initialization phase, system in a mode that measurement is not possible, etc.)*)
    bds_inCmn_notAvl_E,
	(*Not available due to an internal error (e.g., ADC broken)*)
    bds_inCmn_errInt_E,
	(*Precondition is not met*)
    bds_inCmn_invldCfg_E,
	(*API call invalid (e.g., configuration invalid for the requested signal, etc.)*)
    bds_inCmn_invldPrm_E,
	(*API call invalid (e.g., incorrect parameters, etc.)*)
    bds_inCmn_errPrecon_E
)USINT;
END_TYPE

// I/O API/IN/ENUM/bds_inCmn_pullType_te
(*Enumeration of the pull status option.*)
{attribute 'external_name' := 'cmp_rts_bds_inCmn_pullType_te'}
TYPE bds_inCmn_pullType_te :
(
	(*Pull up to 5V*)
    bds_inCmn_pull5V_E :=0,
	(*Pull up to UBatt*)
    bds_inCmn_pullUbatt_E,
	(*Pull down*)
    bds_inCmn_pullDown_E,
	(*External*)
    bds_inCmn_pullExternal_E,
	(*Number of possible pull type selection*)
    bds_inCmn_pullType_num_E
)USINT;
END_TYPE

// I/O API/IN/ENUM/bds_inI_stShunt_te
(*Enumeration encoding the status of an input shunt resistor used for current measurement.*)
{attribute 'external_name' := 'cmp_rts_bds_inI_stShunt_te'}
TYPE bds_inI_stShunt_te :
(
	(*Shunt for current measurement is deactivated*)
    bds_inI_shuntOff_E :=0,
	(*Shunt for current measurement is activated*)
    bds_inI_shuntOn_E,
	(*Overcurrent detected and shunt for current measurement is deactivated*)
    bds_inI_shuntOverCur_E
)USINT;
END_TYPE

// I/O API/IN/ENUM/bds_inCmn_iPull_te
(*Enumeration of the pull current strength options.*)
{attribute 'external_name' := 'cmp_rts_bds_inCmn_iPull_te'}
TYPE bds_inCmn_iPull_te :
(
	(*Current strength 7.5 uA for pull up*)
    bds_inCmn_iPullUp_7_5uA_E :=0,
	(*Current strength 20 uA for pull up and pull down*)
    bds_inCmn_iPull_20uA_E,
	(*Current strength 100 uA for pull down*)
    bds_inCmn_iPullDown_100uA_E,
	(*Current strength 250 uA for pull up*)
    bds_inCmn_iPullUp_250uA_E,
	(*Current strength 500 uA for pull up and pull down*)
    bds_inCmn_iPull_500uA_E,
	(*Current strength 600 uA for pull down*)
    bds_inCmn_iPullDown_600uA_E,
	(*Current strength 1 mA for pull up and pull down*)
    bds_inCmn_iPull_1mA_E,
	(*Current strength  5 mA for pull up and pull down *)
    bds_inCmn_iPull_5mA_E,
	(*Current strength 10 mA for pull up and pull down*)
    bds_inCmn_iPull_10mA_E,
	(*Current strength 20 mA for pull up and pull down *)
    bds_inCmn_iPull_20mA_E,
	(*Restore to default value set by easyConfig *)
    bds_inCmn_iPull_default_E,
	(*Do not change the current strength*)
    bds_inCmn_iPull_noChg_E,
	(*Number of possible current strength selection*)
    bds_inCmn_iPull_num_E
)USINT;
END_TYPE

// I/O API/IN/STRUCTURE/bds_inPwm_tiMeasmt_ts
(*Data structure for one pwm measurement value of the API function |bds_inPwm_getTi|.*)
{attribute 'external_name' := 'cmp_rts_bds_inPwm_tiMeasmt_ts'}
TYPE bds_inPwm_tiMeasmt_ts :
STRUCT
	(*Input period time in [ns]*)
	tiPerd_ns_u32: UDINT;
	(*Input ON time of period in [ns]*)
	tiOnWidth_ns_u32: UDINT;
	(*Number of pulses received (15 bit counter)*)
	cntPls_u32: UDINT;
	(*Status of the measurement*)
	status_e: bds_inCmn_status_te;	
END_STRUCT
END_TYPE

// I/O API/IN/STRUCTURE/bds_inPwm_tiBufdMeasmt_ts
(*Data structure for twenty pwm measurement values of the API function |bds_inPwm_getTiBufd|, used to get the buffered values.*)
{attribute 'external_name' := 'cmp_rts_bds_inPwm_tiBufdMeasmt_ts'}
TYPE bds_inPwm_tiBufdMeasmt_ts :
STRUCT
	(*Up to 20 samples of PWM period in ns, 0th index is latest*)
	tiPerd_ns_au32: ARRAY[0..19] OF UDINT;
	(*Up to 20 samples of ON pulse width in ns*)
	tiOnWidth_ns_au32: ARRAY[0..19] OF UDINT;
	(*Number of new samples (pulses) received since the last call of API. It is limited to 20 samples.*)
	cntNewSample_u8: USINT;
END_STRUCT
END_TYPE

// I/O API/IN/STRUCTURE/bds_inPwm_frqMeasmt_ts
(*Data structure for one pwm frequency measurement value of the API function |bds_inPwm_getFrq|.*)
{attribute 'external_name' := 'cmp_rts_bds_inPwm_frqMeasmt_ts'}
TYPE bds_inPwm_frqMeasmt_ts :
STRUCT
	(*Value of input frequency in (0.1 Hz)*)
	frq_dHz_u32: UDINT;
	(*Value of duty cycle in permil*)
	dutyCyc_perml_u16: UINT;
	(*Number of pulses received (15 bit counter)*)
	cntPls_u32: UDINT;
	(*Status of the measurement*)
	status_e: bds_inCmn_status_te;	
END_STRUCT
END_TYPE

// I/O API/IN/STRUCTURE/bds_inPwm_tiBufd_ts
(*Data structure for pwm measurement value of the API function |bds_inPwm_getTiBufd|.*)
{attribute 'external_name' := 'cmp_rts_bds_inPwm_tiBufd_ts'}
TYPE bds_inPwm_tiBufd_ts :
STRUCT
	(*Status of the measurement*)
	status_e: bds_inCmn_status_te;	
END_STRUCT
END_TYPE

// I/O API/IN/STRUCTURE/bds_inR_measmt_ts
(*Data structure for one resistance measurement value of the API function |bds_inR_get|.*)
{attribute 'external_name' := 'cmp_rts_bds_inR_measmt_ts'}
TYPE bds_inR_measmt_ts :
STRUCT
	(*Status of the measurement*)
	status_e: bds_inCmn_status_te;
	(*Value of input in ohms*)
	r_ohm_u32: UDINT;	
END_STRUCT
END_TYPE

// I/O API/IN/STRUCTURE/bds_inU_measmt_ts
(*Data structure for one voltage measurement value of the API function |bds_inU_get|.*)
{attribute 'external_name' := 'cmp_rts_bds_inU_measmt_ts'}
TYPE bds_inU_measmt_ts :
STRUCT
	(*Status of the measurement*)
	status_e: bds_inCmn_status_te;
	(*Value of input in mV*)
	u_mV_u16: UINT;	
END_STRUCT
END_TYPE

// I/O API/IN/STRUCTURE/bds_inU_cfgPull_ts
(*Return structure for the API function |bds_inU_cfgPull|.*)
{attribute 'external_name' := 'cmp_rts_bds_inU_cfgPull_ts'}
TYPE bds_inU_cfgPull_ts :
STRUCT
	(*Status of the API call*)
	status_e: bds_inCmn_status_te;
END_STRUCT
END_TYPE

// Communication API/ISOBUS/STRUCTURE/bds_isobus_aperiodicDataboxNum_ts
{attribute 'external_name' := 'cmp_rts_bds_isobus_aperiodicDataboxNum_ts'}
TYPE bds_isobus_aperiodicDataboxNum_ts :
STRUCT
	bufferStrt_s16: INT;
	bufferEnd_s16: INT;
END_STRUCT
END_TYPE

// Communication API/ISOBUS/STRUCTURE/bds_isobus_periodicDataboxNum_ts
{attribute 'external_name' := 'cmp_rts_bds_isobus_periodicDataboxNum_ts'}
TYPE bds_isobus_periodicDataboxNum_ts :
STRUCT
	databoxNum_u16: UINT;
END_STRUCT
END_TYPE

// System API/SYS/STRUCTURE/bds_sys_retValApplSwName_ts
{attribute 'external_name' := 'cmp_rts_bds_sys_retValApplSwName_ts'}
(*Return data structure for |bds_sys_applSwName| API.*)
TYPE bds_sys_retValApplSwName_ts :
STRUCT
	(*Function call status return value.*)  
	status_e : bds_sys_aswNameStatus_te;
END_STRUCT
END_TYPE

// System API/SYS/ENUM/bds_sys_aswNameStatus_te
{attribute 'external_name' := 'cmp_rts_bds_sys_aswNameStatus_te'}
(*Listed all the enumeration return types for |bds_sys_applSwName| function.*)
TYPE bds_sys_aswNameStatus_te :
(
	(*Function is called without errors.*)
    bds_sys_swnmOk_E := 0,
	(*String length of ASW name is too long / invalid parameter.*)
    bds_sys_errSwnm_E
);
END_TYPE

// I/O API/OUT/STRUCTURE/bds_outClcU_setVoltage_ts
{attribute 'external_name' := 'cmp_rts_bds_outClcU_setVoltage_ts'}
TYPE bds_outClcU_setVoltage_ts :
STRUCT
	///
    /// bds_outCmn_ok_E  		API call is successful, signal is valid
    /// bds_outCmn_outOfRng_E 	Requested set voltage has exceeded maximum limit for the signal
    /// bds_outCmn_errInt_E 	API call can not be processed due to an error returned from internal function call
    /// bds_outCmn_errLockd_E 	API call can not be processed, because output is locked
    /// bds_outCmn_invldPrm_E 	API call can not be processed, signal is not configured as ClcU output
	///
	/// Valid only FOR API FUNCTION bds_outClcU_setVoltage_ffi
	///
    /// bds_sentCmn_errFfi_E 	API call can not be processed, FFI access denied
 

	statusApi_e: bds_outCmn_statusApi_te;
END_STRUCT
END_TYPE

// I/O API/OUT/ENUM/bds_outCmn_statusApi_te
{attribute 'external_name' := 'cmp_rts_bds_outCmn_statusApi_te'}
TYPE bds_outCmn_statusApi_te :
(
	bds_outCmn_ok_E := 0,
	bds_outCmn_outOfRng_E := 1,
	bds_outCmn_notAvl_E := 2,
	bds_outCmn_errExt_E := 3,
	bds_outCmn_errInt_E := 4,
	bds_outCmn_errLockd_E := 5,
	bds_outCmn_errDiOutp_E := 6,
	bds_outCmn_invldCfg_E := 7,
	bds_outCmn_invldPrm_E := 8,
	bds_outCmn_errFfi_E := 9
)USINT;
END_TYPE

// I/O API/OUT/STRUCTURE/bds_outClcU_setPercUBat_ts
{attribute 'external_name' := 'cmp_rts_bds_outClcU_setPercUBat_ts'}
TYPE bds_outClcU_setPercUBat_ts :
STRUCT
	///
    /// bds_outCmn_ok_E  		API call is successful, signal is valid
    /// bds_outCmn_outOfRng_E 	Requested set voltage has exceeded maximum limit for the signal
    /// bds_outCmn_errInt_E 	API call can not be processed due to an error returned from internal function call
    /// bds_outCmn_errLockd_E 	API call can not be processed, because output is locked
    /// bds_outCmn_invldPrm_E 	API call can not be processed, signal is not configured as ClcU output
	///
	/// Valid only FOR API FUNCTION bds_outClcU_setVoltage_ffi
	///
    /// bds_sentCmn_errFfi_E 	API call can not be processed, FFI access denied
 

	statusApi_e: bds_outCmn_statusApi_te;
END_STRUCT
END_TYPE

// I/O API/OUT/STRUCTURE/bds_outClcU_get_ts
{attribute 'external_name' := 'cmp_rts_bds_outClcU_get_ts'}
TYPE bds_outClcU_get_ts :
STRUCT
	///
    /// uAct_mV_u16  		    Actual voltage measurement value in [mV]
    /// uSet_mV_u16 	        Current setpoint voltage in [mV]
    /// statusDiag_b 	        Detailed diagnostic information of the ClcU output pin
    /// statusApi_e 	        Status of the BDS function call
 
	uAct_mV_u16: UINT;
	uSet_mV_u16: UINT;
	statusDiag_b: bds_outCmn_statusDiag_tb;
	statusApi_e: bds_outCmn_statusApi_te;
END_STRUCT
END_TYPE

// I/O API/OUT/STRUCTURE/bds_outCmn_statusDiag_tb
(*Bit field type definition for the output module with diagnostic status information of output pin.*)
{attribute 'external_name' := 'cmp_rts_bds_outCmn_statusDiag_tb'}
/// stErrSCB_b1 Fault error status for short cut to battery
/// stErrSCG_b1 :  Fault error status for short cut to ground
/// stErrOL_b1 : Fault error status for open load
///stErrOT_b1 : Fault error status for over temperature
///stErrOC_b1 : Fault error status for over current
/// stErrOR_b1 : Fault error status for out of range
///stUnintdSwtOn_b1 : Status of output pin with unintended switch ON error
/// stLckdByINH_b1 : Status of output pin is locked by inhibit functionality
/// stLckdByHwMon_b1 : Status of output pin is locked by hardware monitoring functionality
/// stDiOutp_b1 : Status of output pin; TRUE: Output is disabled, FALSE: Output is enabled
/// stDiFulDiag_b1 : Status of output pin; TRUE: Full diagnosis is disabled, FALSE: Full diagnosis is enabled
/// stDiOpenLoadDetn_b1 : Status of output pin; TRUE: Open load detection disabled, FALSE: Open Load Detection enabled
/// stDiNonHotSCDetn_b1 : Status of output pin; TRUE: NON-Hot error detection is disabled, FALSE: NON-Hot error detection is enabled
/// stReacvnTmrNotElapsed_b1 : Status wait time of output pin; TRUE: Time for reactivation after hot error short circuit error not elapsed, FALSE: Time for reactivation after hot error short circuit error is elapsed
///resd1_b: unused bits
 

TYPE bds_outCmn_statusDiag_tb :
STRUCT
	stErrSCB_b1: BIT;
	stErrSCG_b1: BIT;
	stErrOL_b1: BIT;
	stErrOT_b1: BIT;
	stErrOC_b1: BIT;
	stErrOR_b1: BIT;
	stUnintdSwtOn_b1: BIT;
	stLckdByINH_b1: BIT;
	stLckdByHwMon_b1: BIT;
	stDiOutp_b1: BIT;
	stDiFulDiag_b1: BIT;
	stDiOpenLoadDetn_b1: BIT;
	stDiNonHotSCDetn_b1: BIT;
	stReacvnTmrNotElapsed_b1: BIT;
	resd1_b: BIT;
END_STRUCT
END_TYPE

// I/O API/OUT/STRUCTURE/bds_outClcU_rstErr_ts
{attribute 'external_name' := 'cmp_rts_bds_outClcU_rstErr_ts'}
TYPE bds_outClcU_rstErr_ts :
STRUCT
	///
    /// statusApi_e 	        Status of the BDS function call
 
	statusApi_e: bds_outCmn_statusApi_te;
END_STRUCT
END_TYPE

// I/O API/OUT/STRUCTURE/bds_outDig_set_ts
{attribute 'external_name' := 'cmp_rts_bds_outDig_set_ts'}
TYPE bds_outDig_set_ts :
STRUCT
	///
    /// statusApi_e 	        Status of the BDS function call
 
	statusApi_e: bds_outCmn_statusApi_te;
END_STRUCT
END_TYPE

// I/O API/OUT/STRUCTURE/bds_outDig_get_ts
{attribute 'external_name' := 'cmp_rts_bds_outDig_get_ts'}
TYPE bds_outDig_get_ts :
STRUCT
	///
	/// Digital status of the selected digital output pin (FALSE = Low/Off, TRUE = High/On)
	stFlgEna_l: BOOL;
	/// Measured current of the selected digital output pin in [mA]
	iAct_mA_u16: UINT;
	/// Bit status information of the selected digital output pin
	statusDiag_b: bds_outCmn_statusDiag_tb;
    /// statusApi_e 	        Status of the BDS function call
 
	statusApi_e: bds_outCmn_statusApi_te;
END_STRUCT
END_TYPE

// I/O API/OUT/STRUCTURE/bds_outDig_cfgDiag_ts
{attribute 'external_name' := 'cmp_rts_bds_outDig_cfgDiag_ts'}
TYPE bds_outDig_cfgDiag_ts :
STRUCT
	///
    /// statusApi_e 	        Status of the BDS function call
 
	statusApi_e: bds_outCmn_statusApi_te;
END_STRUCT
END_TYPE

// I/O API/OUT/STRUCTURE/bds_outDig_rstErr_ts
{attribute 'external_name' := 'cmp_rts_bds_outDig_rstErr_ts'}
TYPE bds_outDig_rstErr_ts :
STRUCT
	///
    /// statusApi_e 	        Status of the BDS function call
 
	statusApi_e: bds_outCmn_statusApi_te;
END_STRUCT
END_TYPE

// I/O API/OUT/STRUCTURE/bds_outPwm_setDutyCycle_ts
{attribute 'external_name' := 'cmp_rts_bds_outPwm_setDutyCycle_ts'}
TYPE bds_outPwm_setDutyCycle_ts :
STRUCT
	///
    /// statusApi_e 	        Status of the BDS function call
 
	statusApi_e: bds_outCmn_statusApi_te;
END_STRUCT
END_TYPE

// I/O API/OUT/STRUCTURE/bds_outPwm_get_ts
{attribute 'external_name' := 'cmp_rtsbds_outPwm_get_ts'}
TYPE bds_outPwm_get_ts :
STRUCT
	///
	/// Setpoint current value in [mA]
	iSet_u16: UINT;
	/// Measured current of the selected digital output pin in [mA]
	iAct_mA_u16: UINT;
	/// Current duty cycle in [permil]
	ratDutyCycle_permil_u16: UINT;
	/// Bit status information of the selected digital output pin
	statusDiag_b: bds_outCmn_statusDiag_tb;
    /// statusApi_e 	        Status of the BDS function call
 
	statusApi_e: bds_outCmn_statusApi_te;
END_STRUCT
END_TYPE

// I/O API/OUT/STRUCTURE/bds_outPwm_cfgPeriod_ts
{attribute 'external_name' := 'cmp_rts_bds_outPwm_cfgPeriod_ts'}
TYPE bds_outPwm_cfgPeriod_ts :
STRUCT
	///
    /// statusApi_e 	        Status of the BDS function call
 
	statusApi_e: bds_outCmn_statusApi_te;
END_STRUCT
END_TYPE

// I/O API/OUT/STRUCTURE/bds_outPwm_rstErr_ts
{attribute 'external_name' := 'cmp_rts_bds_outPwm_rstErr_ts'}
TYPE bds_outPwm_rstErr_ts :
STRUCT
	///
    /// statusApi_e 	        Status of the BDS function call
 
	statusApi_e: bds_outCmn_statusApi_te;
END_STRUCT
END_TYPE

// I/O API/OUT/STRUCTURE/bds_outPwm_cfgDiag_ts
{attribute 'external_name' := 'cmp_rts_bds_outPwm_cfgDiag_ts'}
TYPE bds_outPwm_cfgDiag_ts :
STRUCT
	///
    /// statusApi_e 	        Status of the BDS function call
 
	statusApi_e: bds_outCmn_statusApi_te;
END_STRUCT
END_TYPE

// I/O API/OUT/STRUCTURE/bds_outPwm_cfgMode_ts
{attribute 'external_name' := 'cmp_rts_bds_outPwm_cfgMode_ts'}
TYPE bds_outPwm_cfgMode_ts :
STRUCT
	///
    /// statusApi_e 	        Status of the BDS function call
 
	statusApi_e: bds_outCmn_statusApi_te;
END_STRUCT
END_TYPE

// I/O API/OUT/STRUCTURE/bds_outPwm_setCurrent_ts
{attribute 'external_name' := 'cmp_rts_bds_outPwm_setCurrent_ts'}
TYPE bds_outPwm_setCurrent_ts :
STRUCT
	///
    /// statusApi_e 	        Status of the BDS function call
 
	statusApi_e: bds_outCmn_statusApi_te;
END_STRUCT
END_TYPE

// I/O API/OUT/STRUCTURE/bds_outPwm_cfgDiagCurrentDe_ts
{attribute 'external_name' := 'cmp_rts_bds_outPwm_cfgDiagCurrentDe_ts'}
TYPE bds_outPwm_cfgDiagCurrentDe_ts :
STRUCT
	///
    /// statusApi_e 	        Status of the BDS function call
 
	statusApi_e: bds_outCmn_statusApi_te;
END_STRUCT
END_TYPE

// I/O API/OUT/STRUCTURE/bds_outPwm_cfgDither_ts
{attribute 'external_name' := 'cmp_rts_bds_outPwm_cfgDither_ts'}
TYPE bds_outPwm_cfgDither_ts :
STRUCT
	///
    /// statusApi_e 	        Status of the BDS function call
 
	statusApi_e: bds_outCmn_statusApi_te;
END_STRUCT
END_TYPE

// I/O API/OUT/STRUCTURE/bds_outClcU_cfgClc_ts
{attribute 'external_name' := 'cmp_rts_bds_outClcU_cfgClc_ts'}
TYPE bds_outClcU_cfgClc_ts :
STRUCT
	///
    /// statusApi_e 	        Status of the BDS function call
 
	statusApi_e: bds_outCmn_statusApi_te;
END_STRUCT
END_TYPE

// I/O API/OUT/STRUCTURE/bds_outClcU_clcParams_ts
{attribute 'external_name' := 'cmp_rts_bds_outClcU_clcParams_ts'}
TYPE bds_outClcU_clcParams_ts :
STRUCT
	///
    /// Kp_u16 	        PI controller proportional factor Kp
    /// Ki_u16 	        PI controller integral factor Ki
	Kp_u16: UINT;
	Ki_u16: UINT;
END_STRUCT
END_TYPE

// I/O API/OUT/STRUCTURE/bds_outCmn_diagParam_ts
{attribute 'external_name' := 'cmp_rts_bds_outCmn_diagParam_ts'}
TYPE bds_outCmn_diagParam_ts :
STRUCT
	///
    /// diFullDiag_l  		Enable or disable the full diagnostic;
	///							TRUE = Disable full diagnostic (test pulses are disabled and no full DGDI diagnosis)
	///   						FALSE = Enable full diagnostic (test pulses are enabled for full DGDI diagnosis)

 
    /// diCntlAndDiag_l 	Disable control and diagnostic of the output;
    ///							TRUE = Disable the output and the diagnosis for this output
    ///							FALSE = Enable the output and the diagnosis for this output
 
    /// diOpenLoadDetn_l 	Disable control and diagnostic of the output;
    ///							TRUE = Disable the output and the diagnosis for this output
    ///							FALSE = Enable the output and the diagnosis for this output
	
	/// diNonHotSCDetn_l 	Disable control and diagnostic of the output;
    ///							TRUE = Disable the output and the diagnosis for this output
    ///							FALSE = Enable the output and the diagnosis for this output
 

	diFullDiag_l: BOOL;
	diCntlAndDiag_l: BOOL;
	diOpenLoadDetn_l: BOOL;
	diNonHotSCDetn_l: BOOL;
END_STRUCT
END_TYPE

// I/O API/OUT/STRUCTURE/bds_outPwm_cfgClc_ts
{attribute 'external_name' := 'cmp_rts_Mbds_outPwm_cfgClc_ts'}
TYPE bds_outPwm_cfgClc_ts :
STRUCT
	///
    /// statusApi_e 	        Status of the BDS function call
 
	statusApi_e: bds_outCmn_statusApi_te;
END_STRUCT
END_TYPE

// I/O API/OUT/STRUCTURE/bds_outPwm_clcParams_ts
{attribute 'external_name' := 'cmp_rts_bds_outPwm_clcParams_ts'}
TYPE bds_outPwm_clcParams_ts :
STRUCT
	///
    /// Kp_u16 	        PI controller proportional factor Kp
    /// Ki_u16 	        PI controller integral factor Ki
	Kp_u16: UINT;
	Ki_u16: UINT;
END_STRUCT
END_TYPE

// I/O API/OUT/STRUCTURE/bds_outPwm_ditherParams_ts
{attribute 'external_name' := 'cmp_rts_bds_outPwm_ditherParams_ts'}
TYPE bds_outPwm_ditherParams_ts :
STRUCT
	///
    /// ditherFrq_Hz_e 	        Dither frequency in [Hz]
    ///  ditherAmp_mA_u16       Dither amplitude in [mA]

	ditherFrq_Hz_e: bds_outPwm_cfgDither_te; 
	ditherAmp_mA_u16: UINT;
END_STRUCT
END_TYPE

// I/O API/OUT/ENUM/bds_outPwm_cfgMode_te
{attribute 'external_name' := 'cmp_rts_bds_outPwm_cfgMode_te'}
TYPE bds_outPwm_cfgMode_te :
(
	///  bds_outMode_PWM_E:            PWM output mode
	/// bds_outMode_CLCC_E:            Closed loop control current mode
	bds_outMode_PWM_E := 0,
	bds_outMode_CLCC_E := 1
)USINT;
END_TYPE

// I/O API/OUT/ENUM/bds_outPwm_cfgDither_te
{attribute 'external_name' := 'cmp_rts_bds_outPwm_cfgDither_te'}

/// bds_outPwm_dither_0_Hz_E        0Hz means dither is disabled
/// bds_outPwm_dither_83_Hz_E       Closed loop control dither frequency in [Hz]
/// bds_outPwm_dither_90_Hz_E       Closed loop control dither frequency in [Hz]
/// bds_outPwm_dither_100_Hz_E      Closed loop control dither frequency in [Hz]
/// bds_outPwm_dither_111_Hz_E      Closed loop control dither frequency in [Hz]
/// bds_outPwm_dither_125_Hz_E      Closed loop control dither frequency in [Hz]
/// bds_outPwm_dither_142_Hz_E      Closed loop control dither frequency in [Hz]
/// bds_outPwm_dither_166_Hz_E      Closed loop control dither frequency in [Hz]
/// bds_outPwm_dither_200_Hz_E      Closed loop control dither frequency in [Hz]
/// bds_outPwm_dither_250_Hz_E      Closed loop control dither frequency in [Hz]
 

TYPE bds_outPwm_cfgDither_te :
(
	bds_outPwm_dither_0_Hz_E := 0,
	bds_outPwm_dither_83_Hz_E := 83,
	bds_outPwm_dither_90_Hz_E := 90,
	bds_outPwm_dither_100_Hz_E := 100,
	bds_outPwm_dither_111_Hz_E := 111,
	bds_outPwm_dither_125_Hz_E := 125,
	bds_outPwm_dither_142_Hz_E := 142,
	bds_outPwm_dither_166_Hz_E := 166,
	bds_outPwm_dither_200_Hz_E := 200,
	bds_outPwm_dither_250_Hz_E := 250
)USINT;
END_TYPE

